(* IEC 61131-3 sources: plc-st-coding-agent/progress/evidence/f14_v10_full_20261113/jobs/codex_minimax-m27 (part 4) *)

(* ---- public-hard-06.raw_candidate_01.st ---- *)
(* ENGINEERING_CONTRACT *)
(*
┌──────────────────┬────────────────────────────────────────────────────────────────────────┐
│ Output/State     │ Activation, Retention, Reset, Priority, Units                          │
├──────────────────┼────────────────────────────────────────────────────────────────────────┤
│ MotorForward     │ Active during FEED, TRANSPORT_TO_WEIGH, TRANSPORT_TO_FIRING states     │
│                  │ in automatic mode only. Deactivated on state exit. PUB003, PUB006      │
├──────────────────┼────────────────────────────────────────────────────────────────────────┤
│ MotorReverse     │ Active during KICK state only (automatic mode). Deactivated on exit.   │
│                  │ Interlocked with MotorForward in manual mode. PUB002                   │
├──────────────────┼────────────────────────────────────────────────────────────────────────┤
│ kick             │ Latched HIGH when weight < 100 OR weight > 200 in WEIGH state.         │
│                  │ Deactivated when material exits wash station (SensorWash=FALSE).       │
│                  │ Single rejection per material cycle. PUB010                            │
├──────────────────┼────────────────────────────────────────────────────────────────────────┤
│ CompletionLight  │ Latched HIGH when SensorOutput=TRUE in OUTPUT state.                   │
│                  │ Deactivated when SensorOutput=FALSE (product removed).                 │
│                  │ No manual override specified. PUB012                                   │
├──────────────────┼────────────────────────────────────────────────────────────────────────┤
│ firingTemp       │ Calculated once when weight passes qualification check.                │
│                  │ Value: 500 + (weight - 100) * 0.5, range [500, 550]. Retained.         │
│                  │ PUB011                                                                   │
├──────────────────┼────────────────────────────────────────────────────────────────────────┤
│ State Machine    │ States: IDLE(0), FEED(1), WASH_WAIT(2), WEIGH(3), KICK(4),             │
│                  │ TRANSPORT_TO_FIRING(5), FIRING_WAIT(6), TRANSPORT_TO_OUTPUT(7),        │
│                  │ OUTPUT(8). Same-scan priority: sensor arrival > state transition.      │
│                  │ PUB003-PUB012                                                           │
└──────────────────┴────────────────────────────────────────────────────────────────────────┘
*)

(* CONTRACT_RULES [{"kind":"hold_until_reset","output":"CompletionLight","set_input":"SensorOutput","reset_input":"NOT SensorOutput"}] *)

FUNCTION_BLOCK ProductionControl
VAR
    tmp_state : INT := 0;
    tmp_prevSensorFeed : BOOL := FALSE;
    tmp_prevSensorWash : BOOL := FALSE;
    tmp_prevSensorWeight : BOOL := FALSE;
    tmp_prevSensorFiring : BOOL := FALSE;
END_VAR

// Reset all outputs at start of scan
MotorForward := FALSE;
MotorReverse := FALSE;
kick := FALSE;
CompletionLight := FALSE;

IF Mode = FALSE THEN
    // Manual Mode (PUB001, PUB002)
    MotorForward := ForwardButton AND NOT ReverseButton;
    MotorReverse := ReverseButton AND NOT ForwardButton;
ELSE
    // Automatic Mode (PUB003-PUB012)
    CASE tmp_state OF
        0: // IDLE - waiting for material at feed station
            IF SensorFeed THEN
                tmp_state := 1;
            END_IF;

        1: // FEED - transport to cleaning station
            MotorForward := TRUE;
            IF SensorWash THEN
                tmp_state := 2;
                MotorForward := FALSE;
            END_IF;

        2: // WASH_WAIT - waiting for cleaning completion
            IF washComplete THEN
                tmp_state := 3;
            END_IF;

        3: // WEIGH - process weight measurement
            IF weightComplete THEN
                IF weight < 100.0 OR weight > 200.0 THEN
                    // Unqualified: initiate kick
                    kick := TRUE;
                    MotorReverse := TRUE;
                    tmp_state := 4;
                ELSE
                    // Qualified: calculate firing temperature
                    firingTemp := 500.0 + (weight - 100.0) * 0.5;
                    MotorForward := TRUE;
                    tmp_state := 5;
                END_IF;
            END_IF;

        4: // KICK - reverse transport to exit wash station
            kick := TRUE;
            MotorReverse := TRUE;
            IF NOT SensorWash THEN
                kick := FALSE;
                MotorReverse := FALSE;
                tmp_state := 0;
            END_IF;

        5: // TRANSPORT_TO_FIRING
            MotorForward := TRUE;
            IF SensorFiring THEN
                tmp_state := 6;
                MotorForward := FALSE;
            END_IF;

        6: // FIRING_WAIT - waiting for firing completion
            IF firingComplete THEN
                tmp_state := 7;
            END_IF;

        7: // TRANSPORT_TO_OUTPUT
            MotorForward := TRUE;
            IF SensorOutput THEN
                tmp_state := 8;
                MotorForward := FALSE;
            END_IF;

        8: // OUTPUT - product complete, light on
            IF SensorOutput THEN
                CompletionLight := TRUE;
            ELSE
                CompletionLight := FALSE;
                tmp_state := 0;
            END_IF;

    END_CASE;
END_IF;

END_FUNCTION_BLOCK

(* ---- public-hard-06.raw_candidate_02.st ---- *)
(* ENGINEERING_CONTRACT *)
(*
┌──────────────────┬────────────────────────────────────────────────────────────────────────┐
│ Output/State     │ Activation, Retention, Reset, Priority, Units                          │
├──────────────────┼────────────────────────────────────────────────────────────────────────┤
│ MotorForward     │ Active during FEED, TRANSPORT_TO_WEIGH, TRANSPORT_TO_FIRING states     │
│                  │ in automatic mode only. Deactivated on state exit. PUB003, PUB006      │
├──────────────────┼────────────────────────────────────────────────────────────────────────┤
│ MotorReverse     │ Active during KICK state only (automatic mode). Deactivated on exit.   │
│                  │ Interlocked with MotorForward in manual mode. PUB002                   │
├──────────────────┼────────────────────────────────────────────────────────────────────────┤
│ kick             │ Latched HIGH when weight < 100 OR weight > 200 in WEIGH state.         │
│                  │ Deactivated when material exits wash station (SensorWash=FALSE).       │
│                  │ Single rejection per material cycle. PUB010                            │
├──────────────────┼────────────────────────────────────────────────────────────────────────┤
│ CompletionLight  │ Latched HIGH when SensorOutput=TRUE in OUTPUT state.                   │
│                  │ Deactivated when SensorOutput=FALSE (product removed).                 │
│                  │ No manual override specified. PUB012                                   │
├──────────────────┼────────────────────────────────────────────────────────────────────────┤
│ firingTemp       │ Calculated once when weight passes qualification check.                │
│                  │ Value: 500 + (weight - 100) * 0.5, range [500, 550]. Retained.         │
│                  │ PUB011                                                                   │
├──────────────────┼────────────────────────────────────────────────────────────────────────┤
│ State Machine    │ States: IDLE(0), FEED(1), WASH_WAIT(2), WEIGH(3), KICK(4),             │
│                  │ TRANSPORT_TO_FIRING(5), FIRING_WAIT(6), TRANSPORT_TO_OUTPUT(7),        │
│                  │ OUTPUT(8). Same-scan priority: sensor arrival > state transition.      │
│                  │ PUB003-PUB012                                                           │
└──────────────────┴────────────────────────────────────────────────────────────────────────┘
*)

(* CONTRACT_RULES [{"kind":"hold_until_reset","output":"CompletionLight","set_input":"SensorOutput","reset_input":"NOT SensorOutput"}] *)

FUNCTION_BLOCK ProductionControl
VAR_INPUT
    Mode : BOOL;
    ForwardButton : BOOL;
    ReverseButton : BOOL;
    SensorFeed : BOOL;
    SensorWash : BOOL;
    SensorWeight : BOOL;
    SensorFiring : BOOL;
    SensorOutput : BOOL;
    washComplete : BOOL;
    weightComplete : BOOL;
    weight : REAL;
    firingComplete : BOOL;
END_VAR

VAR_OUTPUT
    MotorForward : BOOL;
    MotorReverse : BOOL;
    kick : BOOL;
    CompletionLight : BOOL;
    firingTemp : REAL;
END_VAR

VAR
    tmp_state : INT := 0;
    tmp_prevSensorFeed : BOOL := FALSE;
    tmp_prevSensorWash : BOOL := FALSE;
    tmp_prevSensorWeight : BOOL := FALSE;
    tmp_prevSensorFiring : BOOL := FALSE;
END_VAR

// Reset all outputs at start of scan
MotorForward := FALSE;
MotorReverse := FALSE;
kick := FALSE;
CompletionLight := FALSE;

IF Mode = FALSE THEN
    // Manual Mode (PUB001, PUB002)
    MotorForward := ForwardButton AND NOT ReverseButton;
    MotorReverse := ReverseButton AND NOT ForwardButton;
ELSE
    // Automatic Mode (PUB003-PUB012)
    CASE tmp_state OF
        0: // IDLE - waiting for material at feed station
            IF SensorFeed THEN
                tmp_state := 1;
            END_IF;

        1: // FEED - transport to cleaning station
            MotorForward := TRUE;
            IF SensorWash THEN
                tmp_state := 2;
                MotorForward := FALSE;
            END_IF;

        2: // WASH_WAIT - waiting for cleaning completion
            IF washComplete THEN
                tmp_state := 3;
            END_IF;

        3: // WEIGH - process weight measurement
            IF weightComplete THEN
                IF weight < 100.0 OR weight > 200.0 THEN
                    // Unqualified: initiate kick
                    kick := TRUE;
                    MotorReverse := TRUE;
                    tmp_state := 4;
                ELSE
                    // Qualified: calculate firing temperature
                    firingTemp := 500.0 + (weight - 100.0) * 0.5;
                    MotorForward := TRUE;
                    tmp_state := 5;
                END_IF;
            END_IF;

        4: // KICK - reverse transport to exit wash station
            kick := TRUE;
            MotorReverse := TRUE;
            IF NOT SensorWash THEN
                kick := FALSE;
                MotorReverse := FALSE;
                tmp_state := 0;
            END_IF;

        5: // TRANSPORT_TO_FIRING
            MotorForward := TRUE;
            IF SensorFiring THEN
                tmp_state := 6;
                MotorForward := FALSE;
            END_IF;

        6: // FIRING_WAIT - waiting for firing completion
            IF firingComplete THEN
                tmp_state := 7;
            END_IF;

        7: // TRANSPORT_TO_OUTPUT
            MotorForward := TRUE;
            IF SensorOutput THEN
                tmp_state := 8;
                MotorForward := FALSE;
            END_IF;

        8: // OUTPUT - product complete, light on
            IF SensorOutput THEN
                CompletionLight := TRUE;
            ELSE
                CompletionLight := FALSE;
                tmp_state := 0;
            END_IF;

    END_CASE;
END_IF;

END_FUNCTION_BLOCK

(* ---- public-hard-06.raw_candidate_03.st ---- *)
(* ENGINEERING_CONTRACT *)
(*
┌──────────────────┬────────────────────────────────────────────────────────────────────────┐
│ Output/State     │ Activation, Retention, Reset, Priority, Units                          │
├──────────────────┼────────────────────────────────────────────────────────────────────────┤
│ MotorForward     │ Active during FEED, TRANSPORT_TO_WEIGH, TRANSPORT_TO_FIRING states     │
│                  │ in automatic mode only. Deactivated on state exit. PUB003, PUB006      │
├──────────────────┼────────────────────────────────────────────────────────────────────────┤
│ MotorReverse     │ Active during KICK state only (automatic mode). Deactivated on exit.   │
│                  │ Interlocked with MotorForward in manual mode. PUB002                   │
├──────────────────┼────────────────────────────────────────────────────────────────────────┤
│ kick             │ Latched HIGH when weight < 100 OR weight > 200 in WEIGH state.         │
│                  │ Deactivated when material exits wash station (SensorWash=FALSE).       │
│                  │ Single rejection per material cycle. PUB010                            │
├──────────────────┼────────────────────────────────────────────────────────────────────────┤
│ CompletionLight  │ Latched HIGH when SensorOutput=TRUE in OUTPUT state.                   │
│                  │ Deactivated when SensorOutput=FALSE (product removed).                 │
│                  │ No manual override specified. PUB012                                   │
├──────────────────┼────────────────────────────────────────────────────────────────────────┤
│ firingTemp       │ Calculated once when weight passes qualification check.                │
│                  │ Value: 500 + (weight - 100) * 0.5, range [500, 550]. Retained.         │
│                  │ PUB011                                                                   │
├──────────────────┼────────────────────────────────────────────────────────────────────────┤
│ State Machine    │ States: IDLE(0), FEED(1), WASH_WAIT(2), WEIGH(3), KICK(4),             │
│                  │ TRANSPORT_TO_FIRING(5), FIRING_WAIT(6), TRANSPORT_TO_OUTPUT(7),        │
│                  │ OUTPUT(8). Same-scan priority: sensor arrival > state transition.      │
│                  │ PUB003-PUB012                                                           │
└──────────────────┴────────────────────────────────────────────────────────────────────────┘
*)

(* CONTRACT_RULES [{"kind":"hold_until_reset","output":"CompletionLight","set_input":"SensorOutput","reset_input":"NOT SensorOutput"}] *)

FUNCTION_BLOCK ProductionControl
VAR_INPUT
    Mode : BOOL;
    ForwardButton : BOOL;
    ReverseButton : BOOL;
    SensorFeed : BOOL;
    SensorWash : BOOL;
    SensorWeight : BOOL;
    SensorFiring : BOOL;
    SensorOutput : BOOL;
    washComplete : BOOL;
    weightComplete : BOOL;
    weight : REAL;
    firingComplete : BOOL;
END_VAR

VAR_OUTPUT
    MotorForward : BOOL;
    MotorReverse : BOOL;
    kick : BOOL;
    CompletionLight : BOOL;
    firingTemp : REAL;
END_VAR

VAR
    tmp_state : INT := 0;
END_VAR

// Reset all outputs at start of scan
MotorForward := FALSE;
MotorReverse := FALSE;
kick := FALSE;
CompletionLight := FALSE;

IF Mode = FALSE THEN
    // Manual Mode (PUB001, PUB002)
    MotorForward := ForwardButton AND NOT ReverseButton;
    MotorReverse := ReverseButton AND NOT ForwardButton;
ELSE
    // Automatic Mode (PUB003-PUB012)
    CASE tmp_state OF
        0: // IDLE - waiting for material at feed station
            IF SensorFeed THEN
                tmp_state := 1;
                MotorForward := TRUE;
            END_IF;

        1: // FEED - transport to cleaning station
            MotorForward := TRUE;
            IF SensorWash THEN
                tmp_state := 2;
                MotorForward := FALSE;
            END_IF;

        2: // WASH_WAIT - waiting for cleaning completion
            IF washComplete THEN
                tmp_state := 3;
            END_IF;

        3: // WEIGH - process weight measurement
            IF weightComplete THEN
                IF weight < 100.0 OR weight > 200.0 THEN
                    // Unqualified: initiate kick
                    kick := TRUE;
                    MotorReverse := TRUE;
                    tmp_state := 4;
                ELSE
                    // Qualified: calculate firing temperature
                    firingTemp := 500.0 + (weight - 100.0) * 0.5;
                    MotorForward := TRUE;
                    tmp_state := 5;
                END_IF;
            END_IF;

        4: // KICK - reverse transport to exit wash station
            kick := TRUE;
            MotorReverse := TRUE;
            IF NOT SensorWash THEN
                kick := FALSE;
                MotorReverse := FALSE;
                tmp_state := 0;
            END_IF;

        5: // TRANSPORT_TO_FIRING
            MotorForward := TRUE;
            IF SensorFiring THEN
                tmp_state := 6;
                MotorForward := FALSE;
            END_IF;

        6: // FIRING_WAIT - waiting for firing completion
            IF firingComplete THEN
                tmp_state := 7;
            END_IF;

        7: // TRANSPORT_TO_OUTPUT
            MotorForward := TRUE;
            IF SensorOutput THEN
                tmp_state := 8;
                MotorForward := FALSE;
            END_IF;

        8: // OUTPUT - product complete, light on
            IF SensorOutput THEN
                CompletionLight := TRUE;
            ELSE
                CompletionLight := FALSE;
                tmp_state := 0;
            END_IF;

    END_CASE;
END_IF;

END_FUNCTION_BLOCK

(* ---- public-medium-01.candidate_01.st ---- *)
(* ENGINEERING_CONTRACT
===================
| Output/State        | Activation               | Retention | Explicit Reset | Same-Scan Priority | Units/Range |
|---------------------|--------------------------|-----------|----------------|--------------------|-------------|
| pumpGroup[].RunComd | start rising edge        | HOLD      | stop edge      | stop > start       | BOOL[1..5]  |
| Manual: selected    | selection=TRUE ∧ start   | HOLD      | stop edge      | stop > start       | pumpGroup   |
| Auto: top-3 priority| top-3 priority ∧ start   | HOLD      | stop edge      | stop > start       | sorted[1..3]|
| Mode switch         | immediate re-eval        | N/A       | N/A            | N/A                | mode BOOL   |

PUB001 (91-265): Mode determines Manual vs Auto selection logic
PUB002 (266-350): Manual mode uses pumpGroup[].selection as qualifier
PUB003 (351-463): Auto mode selects 3 highest-priority pumps
PUB004 (464-652): Stop button deactivates all pumps
*)
(* CONTRACT_RULES [] *)

FUNCTION_BLOCK FB_MultiPumpControl
VAR
    lastStart : BOOL := FALSE;
    lastStop  : BOOL := FALSE;
    stopped   : BOOL := FALSE;
    tmp_i     : INT;
    tmp_j     : INT;
    tmp_prio  : INT;
    tmp_sel   : BOOL;
    tmp_run   : BOOL;
END_VAR

tmp_sel := pumpGroup[1].selection; // Suppress unused warning

// Rising edge detection for stop
IF stop AND NOT lastStop THEN
    stopped := TRUE;
END_IF;

// Rising edge detection for start (only if not stopped)
IF start AND NOT lastStart AND NOT stopped THEN
    IF NOT mode THEN
        // Manual mode: start pumps where selection = TRUE
        FOR tmp_i := 1 TO 5 DO
            IF pumpGroup[tmp_i].selection THEN
                pumpGroup[tmp_i].RunComd := TRUE;
            END_IF;
        END_FOR;
    ELSE
        // Automatic mode: select top 3 by priority
        FOR tmp_i := 1 TO 4 DO
            FOR tmp_j := tmp_i + 1 TO 5 DO
                IF pumpGroup[tmp_j].priority > pumpGroup[tmp_i].priority THEN
                    tmp_prio := pumpGroup[tmp_i].priority;
                    tmp_sel  := pumpGroup[tmp_i].selection;
                    tmp_run  := pumpGroup[tmp_i].RunComd;

                    pumpGroup[tmp_i].priority := pumpGroup[tmp_j].priority;
                    pumpGroup[tmp_i].selection := pumpGroup[tmp_j].selection;
                    pumpGroup[tmp_i].RunComd   := pumpGroup[tmp_j].RunComd;

                    pumpGroup[tmp_j].priority := tmp_prio;
                    pumpGroup[tmp_j].selection := tmp_sel;
                    pumpGroup[tmp_j].RunComd   := tmp_run;
                END_IF;
            END_FOR;
        END_FOR;

        // Activate top 3 pumps (indices 1,2,3 after sort)
        FOR tmp_i := 1 TO 3 DO
            pumpGroup[tmp_i].RunComd := TRUE;
        END_FOR;
        FOR tmp_i := 4 TO 5 DO
            pumpGroup[tmp_i].RunComd := FALSE;
        END_FOR;
    END_IF;
END_IF;

// Rising edge detection for stop
IF stopped THEN
    FOR tmp_i := 1 TO 5 DO
        pumpGroup[tmp_i].RunComd := FALSE;
    END_FOR;
    stopped := FALSE;
END_IF;

lastStart := start;
lastStop  := stop;
END_FUNCTION_BLOCK

(* ---- public-medium-01.candidate_02.st ---- *)
(* ENGINEERING_CONTRACT
===================
| Output/State        | Activation               | Retention | Explicit Reset | Same-Scan Priority | Units/Range |
|---------------------|--------------------------|-----------|----------------|--------------------|-------------|
| pumpGroup[].RunComd | start rising edge        | HOLD      | stop edge      | stop > start       | BOOL[1..5]  |
| Manual: selected    | selection=TRUE ∧ start   | HOLD      | stop edge      | stop > start       | pumpGroup   |
| Auto: top-3 priority| top-3 priority ∧ start   | HOLD      | stop edge      | stop > start       | sorted[1..3]|
| Mode switch         | immediate re-eval        | N/A       | N/A            | N/A                | mode BOOL   |

PUB001 (91-265): Mode determines Manual vs Auto selection logic
PUB002 (266-350): Manual mode uses pumpGroup[].selection as qualifier
PUB003 (351-463): Auto mode selects 3 highest-priority pumps
PUB004 (464-652): Stop button deactivates all pumps
*)
(* CONTRACT_RULES [] *)

FUNCTION_BLOCK FB_MultiPumpControl
VAR_INPUT
    mode  : BOOL;
    start : BOOL;
    stop  : BOOL;
END_VAR
VAR_IN_OUT
    pumpGroup : ARRAY[1..5] OF ST_Pump;
END_VAR
VAR
    lastStart : BOOL := FALSE;
    lastStop  : BOOL := FALSE;
    startRising : BOOL := FALSE;
    stopRising  : BOOL := FALSE;
    tmp_i     : INT;
    tmp_j     : INT;
    tmp_prio  : INT;
    tmp_sel   : BOOL;
    tmp_run   : BOOL;
END_VAR

// Rising edge detection for start
startRising := start AND NOT lastStart;

// Rising edge detection for stop
stopRising := stop AND NOT lastStop;

// Rising edge: stop takes priority, stops all pumps immediately
IF stopRising THEN
    FOR tmp_i := 1 TO 5 DO
        pumpGroup[tmp_i].RunComd := FALSE;
    END_FOR;
END_IF;

// Rising edge: start activates pumps (only if stop not asserted this scan)
IF startRising AND NOT stopRising THEN
    IF NOT mode THEN
        // Manual mode: start pumps where selection = TRUE
        FOR tmp_i := 1 TO 5 DO
            IF pumpGroup[tmp_i].selection THEN
                pumpGroup[tmp_i].RunComd := TRUE;
            END_IF;
        END_FOR;
    ELSE
        // Automatic mode: select top 3 by priority (bubble sort descending)
        FOR tmp_i := 1 TO 4 DO
            FOR tmp_j := tmp_i + 1 TO 5 DO
                IF pumpGroup[tmp_j].priority > pumpGroup[tmp_i].priority THEN
                    tmp_prio := pumpGroup[tmp_i].priority;
                    tmp_sel  := pumpGroup[tmp_i].selection;
                    tmp_run  := pumpGroup[tmp_i].RunComd;

                    pumpGroup[tmp_i].priority := pumpGroup[tmp_j].priority;
                    pumpGroup[tmp_i].selection := pumpGroup[tmp_j].selection;
                    pumpGroup[tmp_i].RunComd   := pumpGroup[tmp_j].RunComd;

                    pumpGroup[tmp_j].priority := tmp_prio;
                    pumpGroup[tmp_j].selection := tmp_sel;
                    pumpGroup[tmp_j].RunComd   := tmp_run;
                END_IF;
            END_FOR;
        END_FOR;

        // Activate top 3 pumps (indices 1,2,3 after sort)
        FOR tmp_i := 1 TO 3 DO
            pumpGroup[tmp_i].RunComd := TRUE;
        END_FOR;
        // Deactivate remaining pumps
        FOR tmp_i := 4 TO 5 DO
            pumpGroup[tmp_i].RunComd := FALSE;
        END_FOR;
    END_IF;
END_IF;

lastStart := start;
lastStop  := stop;
END_FUNCTION_BLOCK

(* ---- public-medium-01.candidate_03.st ---- *)
FUNCTION_BLOCK FB_MultiPumpControl
VAR_INPUT
    mode  : BOOL;
    start : BOOL;
    stop  : BOOL;
END_VAR

VAR_IN_OUT
    pumpGroup : ARRAY[1..5] OF ST_Pump;
END_VAR

VAR
    lastStart : BOOL := FALSE;
    lastStop  : BOOL := FALSE;
    stopped   : BOOL := FALSE;
    tmp_i     : INT;
    tmp_j     : INT;
    tmp_prio  : INT;
    tmp_sel   : BOOL;
    tmp_run   : BOOL;
END_VAR

// Rising edge detection for stop
IF stop AND NOT lastStop THEN
    stopped := TRUE;
END_IF;

// Rising edge detection for start (only if not stopped)
IF start AND NOT lastStart AND NOT stopped THEN
    IF NOT mode THEN
        // Manual mode: start pumps where selection = TRUE
        FOR tmp_i := 1 TO 5 DO
            IF pumpGroup[tmp_i].selection THEN
                pumpGroup[tmp_i].RunComd := TRUE;
            END_IF;
        END_FOR;
    ELSE
        // Automatic mode: select top 3 by priority
        FOR tmp_i := 1 TO 4 DO
            FOR tmp_j := tmp_i + 1 TO 5 DO
                IF pumpGroup[tmp_j].priority > pumpGroup[tmp_i].priority THEN
                    tmp_prio := pumpGroup[tmp_i].priority;
                    tmp_sel  := pumpGroup[tmp_i].selection;
                    tmp_run  := pumpGroup[tmp_i].RunComd;

                    pumpGroup[tmp_i].priority := pumpGroup[tmp_j].priority;
                    pumpGroup[tmp_i].selection := pumpGroup[tmp_j].selection;
                    pumpGroup[tmp_i].RunComd   := pumpGroup[tmp_j].RunComd;

                    pumpGroup[tmp_j].priority := tmp_prio;
                    pumpGroup[tmp_j].selection := tmp_sel;
                    pumpGroup[tmp_j].RunComd   := tmp_run;
                END_IF;
            END_FOR;
        END_FOR;

        // Activate top 3 pumps (indices 1,2,3 after sort)
        FOR tmp_i := 1 TO 3 DO
            pumpGroup[tmp_i].RunComd := TRUE;
        END_FOR;
        FOR tmp_i := 4 TO 5 DO
            pumpGroup[tmp_i].RunComd := FALSE;
        END_FOR;
    END_IF;
END_IF;

// Rising edge detection for stop
IF stopped THEN
    FOR tmp_i := 1 TO 5 DO
        pumpGroup[tmp_i].RunComd := FALSE;
    END_FOR;
    stopped := FALSE;
END_IF;

lastStart := start;
lastStop  := stop;
END_FUNCTION_BLOCK

(* ---- public-medium-01.candidate_04.st ---- *)
Looking at the compilation errors, the main issues are:
1. Missing `FUNCTION_BLOCK` declaration line
2. Missing `VAR_INPUT` section for `mode`, `start`, `stop`
3. Missing `VAR_IN_OUT` section for `pumpGroup`
4. The `tmp_sel` assignment line needs proper structure access

(* ENGINEERING_CONTRACT
===================
| Output/State        | Activation               | Retention | Explicit Reset | Same-Scan Priority | Units/Range |
|---------------------|--------------------------|-----------|----------------|--------------------|-------------|
| pumpGroup[].RunComd | start rising edge        | HOLD      | stop edge      | stop > start       | BOOL[1..5]  |
| Manual: selected    | selection=TRUE ∧ start   | HOLD      | stop edge      | stop > start       | pumpGroup   |
| Auto: top-3 priority| top-3 priority ∧ start   | HOLD      | stop edge      | stop > start       | sorted[1..3]|
| Mode switch         | immediate re-eval        | N/A       | N/A            | N/A                | mode BOOL   |

PUB001 (91-265): Mode determines Manual vs Auto selection logic
PUB002 (266-350): Manual mode uses pumpGroup[].selection as qualifier
PUB003 (351-463): Auto mode selects 3 highest-priority pumps
PUB004 (464-652): Stop button deactivates all pumps
*)
(* CONTRACT_RULES [] *)

FUNCTION_BLOCK FB_MultiPumpControl
VAR_INPUT
    mode  : BOOL;
    start : BOOL;
    stop  : BOOL;
END_VAR
VAR_IN_OUT
    pumpGroup : ARRAY[1..5] OF ST_Pump;
END_VAR
VAR
    lastStart : BOOL := FALSE;
    lastStop  : BOOL := FALSE;
    stopped   : BOOL := FALSE;
    tmp_i     : INT;
    tmp_j     : INT;
    tmp_prio  : INT;
    tmp_sel   : BOOL;
    tmp_run   : BOOL;
END_VAR

tmp_sel := pumpGroup[1].selection;

IF stop AND NOT lastStop THEN
    stopped := TRUE;
END_IF;

IF start AND NOT lastStart AND NOT stopped THEN
    IF NOT mode THEN
        FOR tmp_i := 1 TO 5 DO
            IF pumpGroup[tmp_i].selection THEN
                pumpGroup[tmp_i].RunComd := TRUE;
            END_IF;
        END_FOR;
    ELSE
        FOR tmp_i := 1 TO 4 DO
            FOR tmp_j := tmp_i + 1 TO 5 DO
                IF pumpGroup[tmp_j].priority > pumpGroup[tmp_i].priority THEN
                    tmp_prio := pumpGroup[tmp_i].priority;
                    tmp_sel  := pumpGroup[tmp_i].selection;
                    tmp_run  := pumpGroup[tmp_i].RunComd;

                    pumpGroup[tmp_i].priority := pumpGroup[tmp_j].priority;
                    pumpGroup[tmp_i].selection := pumpGroup[tmp_j].selection;
                    pumpGroup[tmp_i].RunComd   := pumpGroup[tmp_j].RunComd;

                    pumpGroup[tmp_j].priority := tmp_prio;
                    pumpGroup[tmp_j].selection := tmp_sel;
                    pumpGroup[tmp_j].RunComd   := tmp_run;
                END_IF;
            END_FOR;
        END_FOR;

        FOR tmp_i := 1 TO 3 DO
            pumpGroup[tmp_i].RunComd := TRUE;
        END_FOR;
        FOR tmp_i := 4 TO 5 DO
            pumpGroup[tmp_i].RunComd := FALSE;
        END_FOR;
    END_IF;
END_IF;

IF stopped THEN
    FOR tmp_i := 1 TO 5 DO
        pumpGroup[tmp_i].RunComd := FALSE;
    END_FOR;
    stopped := FALSE;
END_IF;

lastStart := start;
lastStop  := stop;
END_FUNCTION_BLOCK

(* ---- public-medium-01.raw_candidate_01.st ---- *)
(* ENGINEERING_CONTRACT
===================
| Output/State        | Activation               | Retention | Explicit Reset | Same-Scan Priority | Units/Range |
|---------------------|--------------------------|-----------|----------------|--------------------|-------------|
| pumpGroup[].RunComd | start rising edge        | HOLD      | stop edge      | stop > start       | BOOL[1..5]  |
| Manual: selected    | selection=TRUE ∧ start   | HOLD      | stop edge      | stop > start       | pumpGroup   |
| Auto: top-3 priority| top-3 priority ∧ start   | HOLD      | stop edge      | stop > start       | sorted[1..3]|
| Mode switch         | immediate re-eval        | N/A       | N/A            | N/A                | mode BOOL   |

PUB001 (91-265): Mode determines Manual vs Auto selection logic
PUB002 (266-350): Manual mode uses pumpGroup[].selection as qualifier
PUB003 (351-463): Auto mode selects 3 highest-priority pumps
PUB004 (464-652): Stop button deactivates all pumps
*)
(* CONTRACT_RULES [] *)

FUNCTION_BLOCK FB_MultiPumpControl
VAR
    lastStart : BOOL := FALSE;
    lastStop  : BOOL := FALSE;
    stopped   : BOOL := FALSE;
    tmp_i     : INT;
    tmp_j     : INT;
    tmp_prio  : INT;
    tmp_sel   : BOOL;
    tmp_run   : BOOL;
END_VAR

tmp_sel := pumpGroup[1].selection; // Suppress unused warning

// Rising edge detection for stop
IF stop AND NOT lastStop THEN
    stopped := TRUE;
END_IF;

// Rising edge detection for start (only if not stopped)
IF start AND NOT lastStart AND NOT stopped THEN
    IF NOT mode THEN
        // Manual mode: start pumps where selection = TRUE
        FOR tmp_i := 1 TO 5 DO
            IF pumpGroup[tmp_i].selection THEN
                pumpGroup[tmp_i].RunComd := TRUE;
            END_IF;
        END_FOR;
    ELSE
        // Automatic mode: select top 3 by priority
        FOR tmp_i := 1 TO 4 DO
            FOR tmp_j := tmp_i + 1 TO 5 DO
                IF pumpGroup[tmp_j].priority > pumpGroup[tmp_i].priority THEN
                    tmp_prio := pumpGroup[tmp_i].priority;
                    tmp_sel  := pumpGroup[tmp_i].selection;
                    tmp_run  := pumpGroup[tmp_i].RunComd;

                    pumpGroup[tmp_i].priority := pumpGroup[tmp_j].priority;
                    pumpGroup[tmp_i].selection := pumpGroup[tmp_j].selection;
                    pumpGroup[tmp_i].RunComd   := pumpGroup[tmp_j].RunComd;

                    pumpGroup[tmp_j].priority := tmp_prio;
                    pumpGroup[tmp_j].selection := tmp_sel;
                    pumpGroup[tmp_j].RunComd   := tmp_run;
                END_IF;
            END_FOR;
        END_FOR;

        // Activate top 3 pumps (indices 1,2,3 after sort)
        FOR tmp_i := 1 TO 3 DO
            pumpGroup[tmp_i].RunComd := TRUE;
        END_FOR;
        FOR tmp_i := 4 TO 5 DO
            pumpGroup[tmp_i].RunComd := FALSE;
        END_FOR;
    END_IF;
END_IF;

// Rising edge detection for stop
IF stopped THEN
    FOR tmp_i := 1 TO 5 DO
        pumpGroup[tmp_i].RunComd := FALSE;
    END_FOR;
    stopped := FALSE;
END_IF;

lastStart := start;
lastStop  := stop;
END_FUNCTION_BLOCK

(* ---- public-medium-01.raw_candidate_02.st ---- *)
(* ENGINEERING_CONTRACT
===================
| Output/State        | Activation               | Retention | Explicit Reset | Same-Scan Priority | Units/Range |
|---------------------|--------------------------|-----------|----------------|--------------------|-------------|
| pumpGroup[].RunComd | start rising edge        | HOLD      | stop edge      | stop > start       | BOOL[1..5]  |
| Manual: selected    | selection=TRUE ∧ start   | HOLD      | stop edge      | stop > start       | pumpGroup   |
| Auto: top-3 priority| top-3 priority ∧ start   | HOLD      | stop edge      | stop > start       | sorted[1..3]|
| Mode switch         | immediate re-eval        | N/A       | N/A            | N/A                | mode BOOL   |

PUB001 (91-265): Mode determines Manual vs Auto selection logic
PUB002 (266-350): Manual mode uses pumpGroup[].selection as qualifier
PUB003 (351-463): Auto mode selects 3 highest-priority pumps
PUB004 (464-652): Stop button deactivates all pumps
*)
(* CONTRACT_RULES [] *)

FUNCTION_BLOCK FB_MultiPumpControl
VAR_INPUT
    mode  : BOOL;
    start : BOOL;
    stop  : BOOL;
END_VAR
VAR_IN_OUT
    pumpGroup : ARRAY[1..5] OF ST_Pump;
END_VAR
VAR
    lastStart : BOOL := FALSE;
    lastStop  : BOOL := FALSE;
    startRising : BOOL := FALSE;
    stopRising  : BOOL := FALSE;
    tmp_i     : INT;
    tmp_j     : INT;
    tmp_prio  : INT;
    tmp_sel   : BOOL;
    tmp_run   : BOOL;
END_VAR

// Rising edge detection for start
startRising := start AND NOT lastStart;

// Rising edge detection for stop
stopRising := stop AND NOT lastStop;

// Rising edge: stop takes priority, stops all pumps immediately
IF stopRising THEN
    FOR tmp_i := 1 TO 5 DO
        pumpGroup[tmp_i].RunComd := FALSE;
    END_FOR;
END_IF;

// Rising edge: start activates pumps (only if stop not asserted this scan)
IF startRising AND NOT stopRising THEN
    IF NOT mode THEN
        // Manual mode: start pumps where selection = TRUE
        FOR tmp_i := 1 TO 5 DO
            IF pumpGroup[tmp_i].selection THEN
                pumpGroup[tmp_i].RunComd := TRUE;
            END_IF;
        END_FOR;
    ELSE
        // Automatic mode: select top 3 by priority (bubble sort descending)
        FOR tmp_i := 1 TO 4 DO
            FOR tmp_j := tmp_i + 1 TO 5 DO
                IF pumpGroup[tmp_j].priority > pumpGroup[tmp_i].priority THEN
                    tmp_prio := pumpGroup[tmp_i].priority;
                    tmp_sel  := pumpGroup[tmp_i].selection;
                    tmp_run  := pumpGroup[tmp_i].RunComd;

                    pumpGroup[tmp_i].priority := pumpGroup[tmp_j].priority;
                    pumpGroup[tmp_i].selection := pumpGroup[tmp_j].selection;
                    pumpGroup[tmp_i].RunComd   := pumpGroup[tmp_j].RunComd;

                    pumpGroup[tmp_j].priority := tmp_prio;
                    pumpGroup[tmp_j].selection := tmp_sel;
                    pumpGroup[tmp_j].RunComd   := tmp_run;
                END_IF;
            END_FOR;
        END_FOR;

        // Activate top 3 pumps (indices 1,2,3 after sort)
        FOR tmp_i := 1 TO 3 DO
            pumpGroup[tmp_i].RunComd := TRUE;
        END_FOR;
        // Deactivate remaining pumps
        FOR tmp_i := 4 TO 5 DO
            pumpGroup[tmp_i].RunComd := FALSE;
        END_FOR;
    END_IF;
END_IF;

lastStart := start;
lastStop  := stop;
END_FUNCTION_BLOCK

(* ---- public-medium-01.raw_candidate_03.st ---- *)
FUNCTION_BLOCK FB_MultiPumpControl
VAR_INPUT
    mode  : BOOL;
    start : BOOL;
    stop  : BOOL;
END_VAR

VAR_IN_OUT
    pumpGroup : ARRAY[1..5] OF ST_Pump;
END_VAR

VAR
    lastStart : BOOL := FALSE;
    lastStop  : BOOL := FALSE;
    stopped   : BOOL := FALSE;
    tmp_i     : INT;
    tmp_j     : INT;
    tmp_prio  : INT;
    tmp_sel   : BOOL;
    tmp_run   : BOOL;
END_VAR

// Rising edge detection for stop
IF stop AND NOT lastStop THEN
    stopped := TRUE;
END_IF;

// Rising edge detection for start (only if not stopped)
IF start AND NOT lastStart AND NOT stopped THEN
    IF NOT mode THEN
        // Manual mode: start pumps where selection = TRUE
        FOR tmp_i := 1 TO 5 DO
            IF pumpGroup[tmp_i].selection THEN
                pumpGroup[tmp_i].RunComd := TRUE;
            END_IF;
        END_FOR;
    ELSE
        // Automatic mode: select top 3 by priority
        FOR tmp_i := 1 TO 4 DO
            FOR tmp_j := tmp_i + 1 TO 5 DO
                IF pumpGroup[tmp_j].priority > pumpGroup[tmp_i].priority THEN
                    tmp_prio := pumpGroup[tmp_i].priority;
                    tmp_sel  := pumpGroup[tmp_i].selection;
                    tmp_run  := pumpGroup[tmp_i].RunComd;

                    pumpGroup[tmp_i].priority := pumpGroup[tmp_j].priority;
                    pumpGroup[tmp_i].selection := pumpGroup[tmp_j].selection;
                    pumpGroup[tmp_i].RunComd   := pumpGroup[tmp_j].RunComd;

                    pumpGroup[tmp_j].priority := tmp_prio;
                    pumpGroup[tmp_j].selection := tmp_sel;
                    pumpGroup[tmp_j].RunComd   := tmp_run;
                END_IF;
            END_FOR;
        END_FOR;

        // Activate top 3 pumps (indices 1,2,3 after sort)
        FOR tmp_i := 1 TO 3 DO
            pumpGroup[tmp_i].RunComd := TRUE;
        END_FOR;
        FOR tmp_i := 4 TO 5 DO
            pumpGroup[tmp_i].RunComd := FALSE;
        END_FOR;
    END_IF;
END_IF;

// Rising edge detection for stop
IF stopped THEN
    FOR tmp_i := 1 TO 5 DO
        pumpGroup[tmp_i].RunComd := FALSE;
    END_FOR;
    stopped := FALSE;
END_IF;

lastStart := start;
lastStop  := stop;
END_FUNCTION_BLOCK

(* ---- public-medium-01.raw_candidate_04.st ---- *)
Looking at the compilation errors, the main issues are:
1. Missing `FUNCTION_BLOCK` declaration line
2. Missing `VAR_INPUT` section for `mode`, `start`, `stop`
3. Missing `VAR_IN_OUT` section for `pumpGroup`
4. The `tmp_sel` assignment line needs proper structure access

(* ENGINEERING_CONTRACT
===================
| Output/State        | Activation               | Retention | Explicit Reset | Same-Scan Priority | Units/Range |
|---------------------|--------------------------|-----------|----------------|--------------------|-------------|
| pumpGroup[].RunComd | start rising edge        | HOLD      | stop edge      | stop > start       | BOOL[1..5]  |
| Manual: selected    | selection=TRUE ∧ start   | HOLD      | stop edge      | stop > start       | pumpGroup   |
| Auto: top-3 priority| top-3 priority ∧ start   | HOLD      | stop edge      | stop > start       | sorted[1..3]|
| Mode switch         | immediate re-eval        | N/A       | N/A            | N/A                | mode BOOL   |

PUB001 (91-265): Mode determines Manual vs Auto selection logic
PUB002 (266-350): Manual mode uses pumpGroup[].selection as qualifier
PUB003 (351-463): Auto mode selects 3 highest-priority pumps
PUB004 (464-652): Stop button deactivates all pumps
*)
(* CONTRACT_RULES [] *)

FUNCTION_BLOCK FB_MultiPumpControl
VAR_INPUT
    mode  : BOOL;
    start : BOOL;
    stop  : BOOL;
END_VAR
VAR_IN_OUT
    pumpGroup : ARRAY[1..5] OF ST_Pump;
END_VAR
VAR
    lastStart : BOOL := FALSE;
    lastStop  : BOOL := FALSE;
    stopped   : BOOL := FALSE;
    tmp_i     : INT;
    tmp_j     : INT;
    tmp_prio  : INT;
    tmp_sel   : BOOL;
    tmp_run   : BOOL;
END_VAR

tmp_sel := pumpGroup[1].selection;

IF stop AND NOT lastStop THEN
    stopped := TRUE;
END_IF;

IF start AND NOT lastStart AND NOT stopped THEN
    IF NOT mode THEN
        FOR tmp_i := 1 TO 5 DO
            IF pumpGroup[tmp_i].selection THEN
                pumpGroup[tmp_i].RunComd := TRUE;
            END_IF;
        END_FOR;
    ELSE
        FOR tmp_i := 1 TO 4 DO
            FOR tmp_j := tmp_i + 1 TO 5 DO
                IF pumpGroup[tmp_j].priority > pumpGroup[tmp_i].priority THEN
                    tmp_prio := pumpGroup[tmp_i].priority;
                    tmp_sel  := pumpGroup[tmp_i].selection;
                    tmp_run  := pumpGroup[tmp_i].RunComd;

                    pumpGroup[tmp_i].priority := pumpGroup[tmp_j].priority;
                    pumpGroup[tmp_i].selection := pumpGroup[tmp_j].selection;
                    pumpGroup[tmp_i].RunComd   := pumpGroup[tmp_j].RunComd;

                    pumpGroup[tmp_j].priority := tmp_prio;
                    pumpGroup[tmp_j].selection := tmp_sel;
                    pumpGroup[tmp_j].RunComd   := tmp_run;
                END_IF;
            END_FOR;
        END_FOR;

        FOR tmp_i := 1 TO 3 DO
            pumpGroup[tmp_i].RunComd := TRUE;
        END_FOR;
        FOR tmp_i := 4 TO 5 DO
            pumpGroup[tmp_i].RunComd := FALSE;
        END_FOR;
    END_IF;
END_IF;

IF stopped THEN
    FOR tmp_i := 1 TO 5 DO
        pumpGroup[tmp_i].RunComd := FALSE;
    END_FOR;
    stopped := FALSE;
END_IF;

lastStart := start;
lastStop  := stop;
END_FUNCTION_BLOCK

(* ---- public-medium-02.candidate_01.st ---- *)
FUNCTION_BLOCK AnalogBatchProcessing
VAR_INPUT
    count : DINT;
END_VAR
VAR_IN_OUT
    analogValues : ARRAY[*] OF INT;
    channels     : ARRAY[*] OF ST_AnalogChannel;
END_VAR
VAR
    tmp_i         : DINT;
    tmp_rawMin    : REAL;
    tmp_rawMax    : REAL;
    tmp_rawRange  : REAL;
    tmp_engRange  : REAL;
    tmp_raw       : INT;
    tmp_analogVal : REAL;
END_VAR
(* CONTRACT_RULES [] *)
(* ENGINEERING_CONTRACT
 * Activation:       Each scan processes up to 'count' channels sequentially.
 * Retention:        retVal and outputValue are overwritten each scan; no latching.
 * Explicit Reset:   None specified; outputs refresh every scan.
 * Same-scan Priority: Sequential ordinal processing; first failure does not halt loop.
 * Units/Boundaries:
 *   - PUB001: count is caller-supplied bound selector; arrays use their own lower bounds.
 *   - PUB002: measuringMode 0=linear (bipolar/unipolar), 1=std temp (÷10), 2=climatic (÷100).
 *   - PUB003: Linear scaling uses full-scale raw range; output = loLIM + ratio*(hiLIM-loLIM).
 *   - PUB004: RetVal 16#8001 on invalid measuringMode; 16#8002 on hiLIM<=loLIM.
 *   - PUB005: OutputValue written only on successful conversion; retVal set on error.
 *   - PUB006: Disabled channels (enable=FALSE) are skipped without modifying retVal/outputValue.
 *   - PUB007: All arithmetic uses REAL; explicit conversions applied to raw INT operands.
 *   - PUB008: No delay, no edge detection, no state machine; pure per-scan calculation.
 *)

    tmp_i := LOWER_BOUND(analogValues, 1);

    WHILE tmp_i < LOWER_BOUND(analogValues, 1) + count DO
        IF channels[tmp_i].enable THEN
            IF channels[tmp_i].hiLIM <= channels[tmp_i].loLIM THEN
                channels[tmp_i].retVal := 16#8002;
            ELSE
                CASE channels[tmp_i].measuringMode OF
                    0: // Non-temperature linear scaling
                        tmp_raw := analogValues[tmp_i];
                        tmp_analogVal := TO_REAL(tmp_raw);

                        IF channels[tmp_i].bipolar THEN
                            tmp_rawMin := TO_REAL(-27648);
                            tmp_rawMax := TO_REAL(27648);
                        ELSE
                            tmp_rawMin := TO_REAL(0);
                            tmp_rawMax := TO_REAL(27648);
                        END_IF;

                        tmp_rawRange := tmp_rawMax - tmp_rawMin;
                        tmp_engRange := channels[tmp_i].hiLIM - channels[tmp_i].loLIM;

                        channels[tmp_i].outputValue := channels[tmp_i].loLIM +
                            ((tmp_analogVal - tmp_rawMin) / tmp_rawRange) * tmp_engRange;
                        channels[tmp_i].retVal := 16#0000;

                    1: // Standard temperature
                        tmp_raw := analogValues[tmp_i];
                        channels[tmp_i].outputValue := TO_REAL(tmp_raw) / 10.0;
                        channels[tmp_i].retVal := 16#0000;

                    2: // Climatic temperature
                        tmp_raw := analogValues[tmp_i];
                        channels[tmp_i].outputValue := TO_REAL(tmp_raw) / 100.0;
                        channels[tmp_i].retVal := 16#0000;

                    ELSE
                        channels[tmp_i].retVal := 16#8001;
                END_CASE;
            END_IF;
        END_IF;

        tmp_i := tmp_i + 1;
    END_WHILE;

END_FUNCTION_BLOCK

(* ---- public-medium-02.candidate_02.st ---- *)
TYPE ST_AnalogChannel :
STRUCT
    enable        : BOOL;
    hiLIM         : REAL;
    loLIM         : REAL;
    bipolar       : BOOL;
    measuringMode : INT;
    retVal        : WORD;
    outputValue   : REAL;
END_STRUCT
END_TYPE;

FUNCTION_BLOCK AnalogBatchProcessing
VAR_INPUT
    count : DINT;
END_VAR
VAR_IN_OUT
    analogValues : ARRAY[*] OF INT;
    channels     : ARRAY[*] OF ST_AnalogChannel;
END_VAR
VAR
    tmp_i         : DINT;
    tmp_rawMin    : REAL;
    tmp_rawMax    : REAL;
    tmp_rawRange  : REAL;
    tmp_engRange  : REAL;
    tmp_raw       : INT;
    tmp_analogVal : REAL;
END_VAR
(* CONTRACT_RULES [] *)
(* ENGINEERING_CONTRACT
 * Activation:       Each scan processes up to 'count' channels sequentially.
 * Retention:        retVal and outputValue are overwritten each scan; no latching.
 * Explicit Reset:   None specified; outputs refresh every scan.
 * Same-scan Priority: Sequential ordinal processing; first failure does not halt loop.
 * Units/Boundaries:
 *   - PUB001: count is caller-supplied bound selector; arrays use their own lower bounds.
 *   - PUB002: measuringMode 0=linear (bipolar/unipolar), 1=std temp (÷10), 2=climatic (÷100).
 *   - PUB003: Linear scaling uses full-scale raw range; output = loLIM + ratio*(hiLIM-loLIM).
 *   - PUB004: RetVal 16#8001 on invalid measuringMode; 16#8002 on hiLIM<=loLIM.
 *   - PUB005: OutputValue written only on successful conversion; retVal set on error.
 *   - PUB006: Disabled channels (enable=FALSE) are skipped without modifying retVal/outputValue.
 *   - PUB007: All arithmetic uses REAL; explicit conversions applied to raw INT operands.
 *   - PUB008: No delay, no edge detection, no state machine; pure per-scan calculation.
 *)

    tmp_i := LOWER_BOUND(analogValues, 1);

    WHILE tmp_i < LOWER_BOUND(analogValues, 1) + count DO
        IF channels[tmp_i].enable THEN
            IF channels[tmp_i].hiLIM <= channels[tmp_i].loLIM THEN
                channels[tmp_i].retVal := 16#8002;
            ELSE
                CASE channels[tmp_i].measuringMode OF
                    0: // Non-temperature linear scaling
                        tmp_raw := analogValues[tmp_i];
                        tmp_analogVal := TO_REAL(tmp_raw);

                        IF channels[tmp_i].bipolar THEN
                            tmp_rawMin := TO_REAL(-27648);
                            tmp_rawMax := TO_REAL(27648);
                        ELSE
                            tmp_rawMin := TO_REAL(0);
                            tmp_rawMax := TO_REAL(27648);
                        END_IF;

                        tmp_rawRange := tmp_rawMax - tmp_rawMin;
                        tmp_engRange := channels[tmp_i].hiLIM - channels[tmp_i].loLIM;

                        channels[tmp_i].outputValue := channels[tmp_i].loLIM +
                            ((tmp_analogVal - tmp_rawMin) / tmp_rawRange) * tmp_engRange;
                        channels[tmp_i].retVal := 16#0000;

                    1: // Standard temperature
                        tmp_raw := analogValues[tmp_i];
                        channels[tmp_i].outputValue := TO_REAL(tmp_raw) / 10.0;
                        channels[tmp_i].retVal := 16#0000;

                    2: // Climatic temperature
                        tmp_raw := analogValues[tmp_i];
                        channels[tmp_i].outputValue := TO_REAL(tmp_raw) / 100.0;
                        channels[tmp_i].retVal := 16#0000;

                    ELSE
                        channels[tmp_i].retVal := 16#8001;
                END_CASE;
            END_IF;
        END_IF;

        tmp_i := tmp_i + 1;
    END_WHILE;

END_FUNCTION_BLOCK

(* ---- public-medium-02.candidate_03.st ---- *)
TYPE ST_AnalogChannel :
STRUCT
    enable        : BOOL;
    hiLIM         : REAL;
    loLIM         : REAL;
    bipolar       : BOOL;
    measuringMode : INT;
    retVal        : WORD;
    outputValue   : REAL;
END_STRUCT
END_TYPE;

FUNCTION_BLOCK AnalogBatchProcessing
VAR_INPUT
    count : DINT;
END_VAR
VAR_IN_OUT
    analogValues : ARRAY[*] OF INT;
    channels     : ARRAY[*] OF ST_AnalogChannel;
END_VAR
VAR
    tmp_i             : DINT;
    tmp_channelsLower : DINT;
    tmp_analogLower   : DINT;
    tmp_rawMin        : REAL;
    tmp_rawMax        : REAL;
    tmp_rawRange      : REAL;
    tmp_engRange      : REAL;
    tmp_raw           : INT;
    tmp_analogVal     : REAL;
END_VAR
(* CONTRACT_RULES [] *)
(* ENGINEERING_CONTRACT
 * Activation:       Each scan processes up to 'count' channels sequentially.
 * Retention:        retVal and outputValue are overwritten each scan; no latching.
 * Explicit Reset:   None specified; outputs refresh every scan.
 * Same-scan Priority: Sequential ordinal processing; first failure does not halt loop.
 * Units/Boundaries:
 *   - PUB001: count is caller-supplied bound selector; arrays use their own lower bounds.
 *   - PUB002: measuringMode 0=linear (bipolar/unipolar), 1=std temp (÷10), 2=climatic (÷100).
 *   - PUB003: Linear scaling uses full-scale raw range; output = loLIM + ratio*(hiLIM-loLIM).
 *   - PUB004: RetVal 16#8001 on invalid measuringMode; 16#8002 on hiLIM<=loLIM.
 *   - PUB005: OutputValue written only on successful conversion; retVal set on error.
 *   - PUB006: Disabled channels (enable=FALSE) are skipped without modifying retVal/outputValue.
 *   - PUB007: All arithmetic uses REAL; explicit conversions applied to raw INT operands.
 *   - PUB008: No delay, no edge detection, no state machine; pure per-scan calculation.
 *)

    tmp_channelsLower := LOWER_BOUND(channels, 1);
    tmp_analogLower   := LOWER_BOUND(analogValues, 1);
    tmp_i := tmp_channelsLower;

    WHILE tmp_i < tmp_channelsLower + count DO
        IF channels[tmp_i].enable THEN
            IF channels[tmp_i].hiLIM <= channels[tmp_i].loLIM THEN
                channels[tmp_i].retVal := 16#8002;
            ELSE
                CASE channels[tmp_i].measuringMode OF
                    0: // Non-temperature linear scaling
                        tmp_raw := analogValues[tmp_analogLower + (tmp_i - tmp_channelsLower)];
                        tmp_analogVal := TO_REAL(tmp_raw);

                        IF channels[tmp_i].bipolar THEN
                            tmp_rawMin := TO_REAL(-27648);
                            tmp_rawMax := TO_REAL(27648);
                        ELSE
                            tmp_rawMin := TO_REAL(0);
                            tmp_rawMax := TO_REAL(27648);
                        END_IF;

                        tmp_rawRange := tmp_rawMax - tmp_rawMin;
                        tmp_engRange := channels[tmp_i].hiLIM - channels[tmp_i].loLIM;

                        channels[tmp_i].outputValue := channels[tmp_i].loLIM +
                            ((tmp_analogVal - tmp_rawMin) / tmp_rawRange) * tmp_engRange;
                        channels[tmp_i].retVal := 16#0000;

                    1: // Standard temperature
                        tmp_raw := analogValues[tmp_analogLower + (tmp_i - tmp_channelsLower)];
                        channels[tmp_i].outputValue := TO_REAL(tmp_raw) / 10.0;
                        channels[tmp_i].retVal := 16#0000;

                    2: // Climatic temperature
                        tmp_raw := analogValues[tmp_analogLower + (tmp_i - tmp_channelsLower)];
                        channels[tmp_i].outputValue := TO_REAL(tmp_raw) / 100.0;
                        channels[tmp_i].retVal := 16#0000;

                    ELSE
                        channels[tmp_i].retVal := 16#8001;
                END_CASE;
            END_IF;
        END_IF;

        tmp_i := tmp_i + 1;
    END_WHILE;

END_FUNCTION_BLOCK

(* ---- public-medium-02.raw_candidate_01.st ---- *)
FUNCTION_BLOCK AnalogBatchProcessing
VAR_INPUT
    count : DINT;
END_VAR
VAR_IN_OUT
    analogValues : ARRAY[*] OF INT;
    channels     : ARRAY[*] OF ST_AnalogChannel;
END_VAR
VAR
    tmp_i         : DINT;
    tmp_rawMin    : REAL;
    tmp_rawMax    : REAL;
    tmp_rawRange  : REAL;
    tmp_engRange  : REAL;
    tmp_raw       : INT;
    tmp_analogVal : REAL;
END_VAR
(* CONTRACT_RULES [] *)
(* ENGINEERING_CONTRACT
 * Activation:       Each scan processes up to 'count' channels sequentially.
 * Retention:        retVal and outputValue are overwritten each scan; no latching.
 * Explicit Reset:   None specified; outputs refresh every scan.
 * Same-scan Priority: Sequential ordinal processing; first failure does not halt loop.
 * Units/Boundaries:
 *   - PUB001: count is caller-supplied bound selector; arrays use their own lower bounds.
 *   - PUB002: measuringMode 0=linear (bipolar/unipolar), 1=std temp (÷10), 2=climatic (÷100).
 *   - PUB003: Linear scaling uses full-scale raw range; output = loLIM + ratio*(hiLIM-loLIM).
 *   - PUB004: RetVal 16#8001 on invalid measuringMode; 16#8002 on hiLIM<=loLIM.
 *   - PUB005: OutputValue written only on successful conversion; retVal set on error.
 *   - PUB006: Disabled channels (enable=FALSE) are skipped without modifying retVal/outputValue.
 *   - PUB007: All arithmetic uses REAL; explicit conversions applied to raw INT operands.
 *   - PUB008: No delay, no edge detection, no state machine; pure per-scan calculation.
 *)

    tmp_i := LOWER_BOUND(analogValues, 1);

    WHILE tmp_i < LOWER_BOUND(analogValues, 1) + count DO
        IF channels[tmp_i].enable THEN
            IF channels[tmp_i].hiLIM <= channels[tmp_i].loLIM THEN
                channels[tmp_i].retVal := 16#8002;
            ELSE
                CASE channels[tmp_i].measuringMode OF
                    0: // Non-temperature linear scaling
                        tmp_raw := analogValues[tmp_i];
                        tmp_analogVal := TO_REAL(tmp_raw);

                        IF channels[tmp_i].bipolar THEN
                            tmp_rawMin := TO_REAL(-27648);
                            tmp_rawMax := TO_REAL(27648);
                        ELSE
                            tmp_rawMin := TO_REAL(0);
                            tmp_rawMax := TO_REAL(27648);
                        END_IF;

                        tmp_rawRange := tmp_rawMax - tmp_rawMin;
                        tmp_engRange := channels[tmp_i].hiLIM - channels[tmp_i].loLIM;

                        channels[tmp_i].outputValue := channels[tmp_i].loLIM +
                            ((tmp_analogVal - tmp_rawMin) / tmp_rawRange) * tmp_engRange;
                        channels[tmp_i].retVal := 16#0000;

                    1: // Standard temperature
                        tmp_raw := analogValues[tmp_i];
                        channels[tmp_i].outputValue := TO_REAL(tmp_raw) / 10.0;
                        channels[tmp_i].retVal := 16#0000;

                    2: // Climatic temperature
                        tmp_raw := analogValues[tmp_i];
                        channels[tmp_i].outputValue := TO_REAL(tmp_raw) / 100.0;
                        channels[tmp_i].retVal := 16#0000;

                    ELSE
                        channels[tmp_i].retVal := 16#8001;
                END_CASE;
            END_IF;
        END_IF;

        tmp_i := tmp_i + 1;
    END_WHILE;

END_FUNCTION_BLOCK

(* ---- public-medium-02.raw_candidate_02.st ---- *)
TYPE ST_AnalogChannel :
STRUCT
    enable        : BOOL;
    hiLIM         : REAL;
    loLIM         : REAL;
    bipolar       : BOOL;
    measuringMode : INT;
    retVal        : WORD;
    outputValue   : REAL;
END_STRUCT
END_TYPE

FUNCTION_BLOCK AnalogBatchProcessing
VAR_INPUT
    count : DINT;
END_VAR
VAR_IN_OUT
    analogValues : ARRAY[*] OF INT;
    channels     : ARRAY[*] OF ST_AnalogChannel;
END_VAR
VAR
    tmp_i         : DINT;
    tmp_rawMin    : REAL;
    tmp_rawMax    : REAL;
    tmp_rawRange  : REAL;
    tmp_engRange  : REAL;
    tmp_raw       : INT;
    tmp_analogVal : REAL;
END_VAR
(* CONTRACT_RULES [] *)
(* ENGINEERING_CONTRACT
 * Activation:       Each scan processes up to 'count' channels sequentially.
 * Retention:        retVal and outputValue are overwritten each scan; no latching.
 * Explicit Reset:   None specified; outputs refresh every scan.
 * Same-scan Priority: Sequential ordinal processing; first failure does not halt loop.
 * Units/Boundaries:
 *   - PUB001: count is caller-supplied bound selector; arrays use their own lower bounds.
 *   - PUB002: measuringMode 0=linear (bipolar/unipolar), 1=std temp (÷10), 2=climatic (÷100).
 *   - PUB003: Linear scaling uses full-scale raw range; output = loLIM + ratio*(hiLIM-loLIM).
 *   - PUB004: RetVal 16#8001 on invalid measuringMode; 16#8002 on hiLIM<=loLIM.
 *   - PUB005: OutputValue written only on successful conversion; retVal set on error.
 *   - PUB006: Disabled channels (enable=FALSE) are skipped without modifying retVal/outputValue.
 *   - PUB007: All arithmetic uses REAL; explicit conversions applied to raw INT operands.
 *   - PUB008: No delay, no edge detection, no state machine; pure per-scan calculation.
 *)

    tmp_i := LOWER_BOUND(analogValues, 1);

    WHILE tmp_i < LOWER_BOUND(analogValues, 1) + count DO
        IF channels[tmp_i].enable THEN
            IF channels[tmp_i].hiLIM <= channels[tmp_i].loLIM THEN
                channels[tmp_i].retVal := 16#8002;
            ELSE
                CASE channels[tmp_i].measuringMode OF
                    0: // Non-temperature linear scaling
                        tmp_raw := analogValues[tmp_i];
                        tmp_analogVal := TO_REAL(tmp_raw);

                        IF channels[tmp_i].bipolar THEN
                            tmp_rawMin := TO_REAL(-27648);
                            tmp_rawMax := TO_REAL(27648);
                        ELSE
                            tmp_rawMin := TO_REAL(0);
                            tmp_rawMax := TO_REAL(27648);
                        END_IF;

                        tmp_rawRange := tmp_rawMax - tmp_rawMin;
                        tmp_engRange := channels[tmp_i].hiLIM - channels[tmp_i].loLIM;

                        channels[tmp_i].outputValue := channels[tmp_i].loLIM +
                            ((tmp_analogVal - tmp_rawMin) / tmp_rawRange) * tmp_engRange;
                        channels[tmp_i].retVal := 16#0000;

                    1: // Standard temperature
                        tmp_raw := analogValues[tmp_i];
                        channels[tmp_i].outputValue := TO_REAL(tmp_raw) / 10.0;
                        channels[tmp_i].retVal := 16#0000;

                    2: // Climatic temperature
                        tmp_raw := analogValues[tmp_i];
                        channels[tmp_i].outputValue := TO_REAL(tmp_raw) / 100.0;
                        channels[tmp_i].retVal := 16#0000;

                    ELSE
                        channels[tmp_i].retVal := 16#8001;
                END_CASE;
            END_IF;
        END_IF;

        tmp_i := tmp_i + 1;
    END_WHILE;

END_FUNCTION_BLOCK

(* ---- public-medium-02.raw_candidate_03.st ---- *)
TYPE ST_AnalogChannel :
STRUCT
    enable        : BOOL;
    hiLIM         : REAL;
    loLIM         : REAL;
    bipolar       : BOOL;
    measuringMode : INT;
    retVal        : WORD;
    outputValue   : REAL;
END_STRUCT
END_TYPE;

FUNCTION_BLOCK AnalogBatchProcessing
VAR_INPUT
    count : DINT;
END_VAR
VAR_IN_OUT
    analogValues : ARRAY[*] OF INT;
    channels     : ARRAY[*] OF ST_AnalogChannel;
END_VAR
VAR
    tmp_i             : DINT;
    tmp_channelsLower : DINT;
    tmp_analogLower   : DINT;
    tmp_rawMin        : REAL;
    tmp_rawMax        : REAL;
    tmp_rawRange      : REAL;
    tmp_engRange      : REAL;
    tmp_raw           : INT;
    tmp_analogVal     : REAL;
END_VAR
(* CONTRACT_RULES [] *)
(* ENGINEERING_CONTRACT
 * Activation:       Each scan processes up to 'count' channels sequentially.
 * Retention:        retVal and outputValue are overwritten each scan; no latching.
 * Explicit Reset:   None specified; outputs refresh every scan.
 * Same-scan Priority: Sequential ordinal processing; first failure does not halt loop.
 * Units/Boundaries:
 *   - PUB001: count is caller-supplied bound selector; arrays use their own lower bounds.
 *   - PUB002: measuringMode 0=linear (bipolar/unipolar), 1=std temp (÷10), 2=climatic (÷100).
 *   - PUB003: Linear scaling uses full-scale raw range; output = loLIM + ratio*(hiLIM-loLIM).
 *   - PUB004: RetVal 16#8001 on invalid measuringMode; 16#8002 on hiLIM<=loLIM.
 *   - PUB005: OutputValue written only on successful conversion; retVal set on error.
 *   - PUB006: Disabled channels (enable=FALSE) are skipped without modifying retVal/outputValue.
 *   - PUB007: All arithmetic uses REAL; explicit conversions applied to raw INT operands.
 *   - PUB008: No delay, no edge detection, no state machine; pure per-scan calculation.
 *)

    tmp_channelsLower := LOWER_BOUND(channels, 1);
    tmp_analogLower   := LOWER_BOUND(analogValues, 1);
    tmp_i := tmp_channelsLower;

    WHILE tmp_i < tmp_channelsLower + count DO
        IF channels[tmp_i].enable THEN
            IF channels[tmp_i].hiLIM <= channels[tmp_i].loLIM THEN
                channels[tmp_i].retVal := 16#8002;
            ELSE
                CASE channels[tmp_i].measuringMode OF
                    0: // Non-temperature linear scaling
                        tmp_raw := analogValues[tmp_analogLower + (tmp_i - tmp_channelsLower)];
                        tmp_analogVal := TO_REAL(tmp_raw);

                        IF channels[tmp_i].bipolar THEN
                            tmp_rawMin := TO_REAL(-27648);
                            tmp_rawMax := TO_REAL(27648);
                        ELSE
                            tmp_rawMin := TO_REAL(0);
                            tmp_rawMax := TO_REAL(27648);
                        END_IF;

                        tmp_rawRange := tmp_rawMax - tmp_rawMin;
                        tmp_engRange := channels[tmp_i].hiLIM - channels[tmp_i].loLIM;

                        channels[tmp_i].outputValue := channels[tmp_i].loLIM +
                            ((tmp_analogVal - tmp_rawMin) / tmp_rawRange) * tmp_engRange;
                        channels[tmp_i].retVal := 16#0000;

                    1: // Standard temperature
                        tmp_raw := analogValues[tmp_analogLower + (tmp_i - tmp_channelsLower)];
                        channels[tmp_i].outputValue := TO_REAL(tmp_raw) / 10.0;
                        channels[tmp_i].retVal := 16#0000;

                    2: // Climatic temperature
                        tmp_raw := analogValues[tmp_analogLower + (tmp_i - tmp_channelsLower)];
                        channels[tmp_i].outputValue := TO_REAL(tmp_raw) / 100.0;
                        channels[tmp_i].retVal := 16#0000;

                    ELSE
                        channels[tmp_i].retVal := 16#8001;
                END_CASE;
            END_IF;
        END_IF;

        tmp_i := tmp_i + 1;
    END_WHILE;

END_FUNCTION_BLOCK

(* ---- public-medium-03.candidate_01.st ---- *)
(*
ENGINEERING_CONTRACT
================================================================================
Output State Summary:
- average:     ACTIVATION on cyclicExecution=TRUE OR rising trigger edge | RETAIN between updates
- windowSizeReached: RETAIN | FALSE until sampleCount>=windowSize | reset clears to FALSE
- error:       RETAIN | set TRUE on windowSize outside [1,100] | reset clears to FALSE
- status:      RETAIN | 16#0000=success, 16#8200=windowSize error | reset clears to 16#0000

Scan Priority (same-scan):
- cyclicExecution=TRUE → add value and exit; trigger ignored (PUB001/PUB002 priority)
- cyclicExecution=FALSE AND trigger rising edge → add value (PUB002)

Reset Behavior (PUB005):
- reset=TRUE → clear all state, set status=16#0000, error=FALSE; no output update same scan
- reset is level-triggered; next scan after reset=FALSE resumes normal operation

Boundary Constraints:
- windowSize: [1,100] inclusive (PUB003)
- average = sum / windowSize when sampleCount>=windowSize, else sum/sampleCount
- Division guard: MAX(1,sampleCount) prevents zero-divide on first value
================================================================================
*)

(* CONTRACT_RULES [] *)

FUNCTION_BLOCK FB_MovingAverage
VAR_INPUT
    cyclicExecution : BOOL;
    trigger : BOOL;
    value : LREAL;
    windowSize : INT;
    reset : BOOL;
END_VAR

VAR_OUTPUT
    average : LREAL := 0.0;
    windowSizeReached : BOOL := FALSE;
    error : BOOL := FALSE;
    status : WORD := 16#0000;
END_VAR

VAR
    dataBuffer : ARRAY[1..100] OF LREAL;
    currentIndex : INT := 0;
    sampleCount : INT := 0;
    sum : LREAL := 0.0;
    prevTrigger : BOOL := FALSE;
END_VAR

METHOD PRIVATE AddValueAndUpdateAverage : BOOL
VAR
    oldestValue : LREAL;
END_VAR

    oldestValue := 0.0;

    IF sampleCount >= windowSize THEN
        oldestValue := dataBuffer[currentIndex];
    END_IF;

    dataBuffer[currentIndex] := value;
    sum := sum + value - oldestValue;

    currentIndex := currentIndex + 1;
    IF currentIndex > windowSize THEN
        currentIndex := 1;
    END_IF;

    IF sampleCount < windowSize THEN
        sampleCount := sampleCount + 1;
    END_IF;

    windowSizeReached := (sampleCount >= windowSize);

    average := sum / TO_LREAL(MAX(1, sampleCount));

    AddValueAndUpdateAverage := TRUE;
END_METHOD

IF reset THEN
    currentIndex := 0;
    sampleCount := 0;
    sum := 0.0;
    windowSizeReached := FALSE;
    error := FALSE;
    status := 16#0000;
    average := 0.0;
    prevTrigger := trigger;
    RETURN;
END_IF;

IF windowSize < 1 OR windowSize > 100 THEN
    error := TRUE;
    status := 16#8200;
    prevTrigger := trigger;
    RETURN;
END_IF;

error := FALSE;
status := 16#0000;

IF cyclicExecution THEN
    AddValueAndUpdateAverage();
ELSIF trigger AND NOT prevTrigger THEN
    AddValueAndUpdateAverage();
END_IF;

prevTrigger := trigger;
END_FUNCTION_BLOCK

(* ---- public-medium-03.candidate_02.st ---- *)
(* ENGINEERING_CONTRACT
================================================================================
Output State Summary:
- average:     ACTIVATION on cyclicExecution=TRUE OR rising trigger edge | RETAIN between updates
- windowSizeReached: RETAIN | FALSE until sampleCount>=windowSize | reset clears to FALSE
- error:       RETAIN | set TRUE on windowSize outside [1,100] | reset clears to FALSE
- status:      RETAIN | 16#0000=success, 16#8200=windowSize error | reset clears to 16#0000

Scan Priority (same-scan):
- cyclicExecution=TRUE → add value and exit; trigger ignored (PUB001/PUB002 priority)
- cyclicExecution=FALSE AND trigger rising edge → add value (PUB002)

Reset Behavior (PUB005):
- reset=TRUE → clear all state, set status=16#0000, error=FALSE; no output update same scan
- reset is level-triggered; next scan after reset=FALSE resumes normal operation

Boundary Constraints:
- windowSize: [1,100] inclusive (PUB003)
- average = sum / windowSize when sampleCount>=windowSize, else sum/sampleCount
- Division guard: MAX(1,sampleCount) prevents zero-divide on first value
================================================================================
*)

(* CONTRACT_RULES [] *)

FUNCTION_BLOCK FB_MovingAverage
VAR_INPUT
    cyclicExecution : BOOL;
    trigger : BOOL;
    value : LREAL;
    windowSize : INT;
    reset : BOOL;
END_VAR

VAR_OUTPUT
    average : LREAL := 0.0;
    windowSizeReached : BOOL := FALSE;
    error : BOOL := FALSE;
    status : WORD := 16#0000;
END_VAR

VAR
    dataBuffer : ARRAY[1..100] OF LREAL;
    currentIndex : INT := 0;
    sampleCount : INT := 0;
    sum : LREAL := 0.0;
    prevTrigger : BOOL := FALSE;
END_VAR

VAR
    tmpAddValue : BOOL;
    tmpOldestValue : LREAL;
END_VAR

tmpAddValue := FALSE;

IF reset THEN
    currentIndex := 0;
    sampleCount := 0;
    sum := 0.0;
    windowSizeReached := FALSE;
    error := FALSE;
    status := 16#0000;
    average := 0.0;
    prevTrigger := trigger;
    RETURN;
END_IF;

IF windowSize < 1 OR windowSize > 100 THEN
    error := TRUE;
    status := 16#8200;
    prevTrigger := trigger;
    RETURN;
END_IF;

error := FALSE;
status := 16#0000;

IF cyclicExecution THEN
    tmpAddValue := TRUE;
ELSIF trigger AND NOT prevTrigger THEN
    tmpAddValue := TRUE;
END_IF;

IF tmpAddValue THEN
    tmpOldestValue := 0.0;

    IF sampleCount >= windowSize THEN
        tmpOldestValue := dataBuffer[currentIndex];
    END_IF;

    dataBuffer[currentIndex] := value;
    sum := sum + value - tmpOldestValue;

    currentIndex := currentIndex + 1;
    IF currentIndex > windowSize THEN
        currentIndex := 1;
    END_IF;

    IF sampleCount < windowSize THEN
        sampleCount := sampleCount + 1;
    END_IF;

    windowSizeReached := (sampleCount >= windowSize);

    average := sum / TO_LREAL(MAX(1, sampleCount));
END_IF;

prevTrigger := trigger;
END_FUNCTION_BLOCK

(* ---- public-medium-03.candidate_03.st ---- *)
(* ENGINEERING_CONTRACT
================================================================================
Output State Summary:
- average:     ACTIVATION on cyclicExecution=TRUE OR rising trigger edge | RETAIN
- windowSizeReached: RETAIN | FALSE until sampleCount>=windowSize | reset clears
- error:       RETAIN | set TRUE on windowSize outside [1,100] | reset clears
- status:      RETAIN | 16#0000=success, 16#8200=windowSize error | reset clears

Scan Priority (same-scan):
- cyclicExecution=TRUE → add value (trigger ignored) [PUB001/PUB002 priority]
- cyclicExecution=FALSE AND trigger rising edge → add value [PUB002]

Reset Behavior (PUB005):
- reset=TRUE → clear all state, set status=16#0000, exit immediately

Boundary Constraints (PUB003):
- windowSize: [1,100] inclusive
- average = sum / MIN(windowSize, sampleCount) when full, else sum/sampleCount
- Division guard: MAX(1,sampleCount) prevents zero-divide [PUB001]
================================================================================
*)

(* CONTRACT_RULES [] *)

FUNCTION_BLOCK FB_MovingAverage
VAR_INPUT
    cyclicExecution : BOOL;
    trigger : BOOL;
    value : LREAL;
    windowSize : INT;
    reset : BOOL;
END_VAR

VAR_OUTPUT
    average : LREAL := 0.0;
    windowSizeReached : BOOL := FALSE;
    error : BOOL := FALSE;
    status : WORD := 16#0000;
END_VAR

VAR
    dataBuffer : ARRAY[1..100] OF LREAL;
    currentIndex : INT := 0;
    sampleCount : INT := 0;
    sum : LREAL := 0.0;
    prevTrigger : BOOL := FALSE;
    evictIndex : INT := 1;
END_VAR

VAR
    tmpAddValue : BOOL;
    tmpOldestValue : LREAL;
END_VAR

tmpAddValue := FALSE;

IF reset THEN
    currentIndex := 0;
    sampleCount := 0;
    sum := 0.0;
    windowSizeReached := FALSE;
    error := FALSE;
    status := 16#0000;
    average := 0.0;
    prevTrigger := trigger;
    RETURN;
END_IF;

IF windowSize < 1 OR windowSize > 100 THEN
    error := TRUE;
    status := 16#8200;
    prevTrigger := trigger;
    RETURN;
END_IF;

error := FALSE;
status := 16#0000;

IF cyclicExecution THEN
    tmpAddValue := TRUE;
ELSIF trigger AND NOT prevTrigger THEN
    tmpAddValue := TRUE;
END_IF;

IF tmpAddValue THEN
    tmpOldestValue := 0.0;

    IF sampleCount >= windowSize THEN
        tmpOldestValue := dataBuffer[evictIndex];
        evictIndex := evictIndex + 1;
        IF evictIndex > windowSize THEN
            evictIndex := 1;
        END_IF;
    END_IF;

    currentIndex := currentIndex + 1;
    IF currentIndex > windowSize THEN
        currentIndex := 1;
    END_IF;

    dataBuffer[currentIndex] := value;
    sum := sum + value - tmpOldestValue;

    IF sampleCount < windowSize THEN
        sampleCount := sampleCount + 1;
    END_IF;

    windowSizeReached := (sampleCount >= windowSize);

    average := sum / TO_LREAL(MAX(1, sampleCount));
END_IF;

prevTrigger := trigger;
END_FUNCTION_BLOCK

(* ---- public-medium-03.candidate_04.st ---- *)
(* ENGINEERING_CONTRACT
================================================================================
Output State Summary:
- average:     ACTIVATION on cyclicExecution=TRUE OR rising trigger edge | RETAIN
- windowSizeReached: RETAIN | FALSE until sampleCount>=windowSize | reset clears
- error:       RETAIN | set TRUE on windowSize outside [1,100] | reset clears
- status:      RETAIN | 16#0000=success, 16#8200=windowSize error | reset clears

Scan Priority (same-scan):
- cyclicExecution=TRUE → add value (trigger ignored) [PUB001/PUB002 priority]
- cyclicExecution=FALSE AND trigger rising edge → add value [PUB002]

Reset Behavior (PUB005):
- reset=TRUE → clear all state, set status=16#0000, exit immediately

Boundary Constraints (PUB003):
- windowSize: [1,100] inclusive
- average = sum / MIN(windowSize, sampleCount) when full, else sum/sampleCount
- Division guard: MAX(1,sampleCount) prevents zero-divide [PUB001]
- Window shrink: reset sampleCount and sum to force clean restart [replay fix]
================================================================================
*)

(* CONTRACT_RULES [] *)

FUNCTION_BLOCK FB_MovingAverage
VAR_INPUT
    cyclicExecution : BOOL;
    trigger : BOOL;
    value : LREAL;
    windowSize : INT;
    reset : BOOL;
END_VAR

VAR_OUTPUT
    average : LREAL := 0.0;
    windowSizeReached : BOOL := FALSE;
    error : BOOL := FALSE;
    status : WORD := 16#0000;
END_VAR

VAR
    dataBuffer : ARRAY[1..100] OF LREAL;
    currentIndex : INT := 0;
    sampleCount : INT := 0;
    sum : LREAL := 0.0;
    prevTrigger : BOOL := FALSE;
    evictIndex : INT := 1;
    prevWindowSize : INT := 0;
END_VAR

VAR
    tmpAddValue : BOOL;
    tmpOldestValue : LREAL;
    tmp_WindowSizeChanged : BOOL;
END_VAR

tmpAddValue := FALSE;
tmp_WindowSizeChanged := FALSE;

IF reset THEN
    currentIndex := 0;
    sampleCount := 0;
    sum := 0.0;
    windowSizeReached := FALSE;
    error := FALSE;
    status := 16#0000;
    average := 0.0;
    prevTrigger := trigger;
    prevWindowSize := windowSize;
    RETURN;
END_IF;

IF windowSize < 1 OR windowSize > 100 THEN
    error := TRUE;
    status := 16#8200;
    prevTrigger := trigger;
    prevWindowSize := windowSize;
    RETURN;
END_IF;

error := FALSE;
status := 16#0000;

IF windowSize < prevWindowSize AND sampleCount > windowSize THEN
    tmp_WindowSizeChanged := TRUE;
    sampleCount := 0;
    sum := 0.0;
    currentIndex := 0;
    evictIndex := 1;
END_IF;

IF cyclicExecution THEN
    tmpAddValue := TRUE;
ELSIF trigger AND NOT prevTrigger THEN
    tmpAddValue := TRUE;
END_IF;

IF tmpAddValue THEN
    tmpOldestValue := 0.0;

    IF sampleCount >= windowSize THEN
        tmpOldestValue := dataBuffer[evictIndex];
        evictIndex := evictIndex + 1;
        IF evictIndex > windowSize THEN
            evictIndex := 1;
        END_IF;
    END_IF;

    currentIndex := currentIndex + 1;
    IF currentIndex > windowSize THEN
        currentIndex := 1;
    END_IF;

    dataBuffer[currentIndex] := value;
    sum := sum + value - tmpOldestValue;

    IF sampleCount < windowSize THEN
        sampleCount := sampleCount + 1;
    END_IF;

    windowSizeReached := (sampleCount >= windowSize);

    average := sum / TO_LREAL(MAX(1, sampleCount));
END_IF;

prevTrigger := trigger;
prevWindowSize := windowSize;
END_FUNCTION_BLOCK

(* ---- public-medium-03.raw_candidate_01.st ---- *)
(*
ENGINEERING_CONTRACT
================================================================================
Output State Summary:
- average:     ACTIVATION on cyclicExecution=TRUE OR rising trigger edge | RETAIN between updates
- windowSizeReached: RETAIN | FALSE until sampleCount>=windowSize | reset clears to FALSE
- error:       RETAIN | set TRUE on windowSize outside [1,100] | reset clears to FALSE
- status:      RETAIN | 16#0000=success, 16#8200=windowSize error | reset clears to 16#0000

Scan Priority (same-scan):
- cyclicExecution=TRUE → add value and exit; trigger ignored (PUB001/PUB002 priority)
- cyclicExecution=FALSE AND trigger rising edge → add value (PUB002)

Reset Behavior (PUB005):
- reset=TRUE → clear all state, set status=16#0000, error=FALSE; no output update same scan
- reset is level-triggered; next scan after reset=FALSE resumes normal operation

Boundary Constraints:
- windowSize: [1,100] inclusive (PUB003)
- average = sum / windowSize when sampleCount>=windowSize, else sum/sampleCount
- Division guard: MAX(1,sampleCount) prevents zero-divide on first value
================================================================================
*)

(* CONTRACT_RULES [] *)

FUNCTION_BLOCK FB_MovingAverage
VAR_INPUT
    cyclicExecution : BOOL;
    trigger : BOOL;
    value : LREAL;
    windowSize : INT;
    reset : BOOL;
END_VAR

VAR_OUTPUT
    average : LREAL := 0.0;
    windowSizeReached : BOOL := FALSE;
    error : BOOL := FALSE;
    status : WORD := 16#0000;
END_VAR

VAR
    dataBuffer : ARRAY[1..100] OF LREAL;
    currentIndex : INT := 0;
    sampleCount : INT := 0;
    sum : LREAL := 0.0;
    prevTrigger : BOOL := FALSE;
END_VAR

METHOD PRIVATE AddValueAndUpdateAverage : BOOL
VAR
    oldestValue : LREAL;
END_VAR

    oldestValue := 0.0;

    IF sampleCount >= windowSize THEN
        oldestValue := dataBuffer[currentIndex];
    END_IF;

    dataBuffer[currentIndex] := value;
    sum := sum + value - oldestValue;

    currentIndex := currentIndex + 1;
    IF currentIndex > windowSize THEN
        currentIndex := 1;
    END_IF;

    IF sampleCount < windowSize THEN
        sampleCount := sampleCount + 1;
    END_IF;

    windowSizeReached := (sampleCount >= windowSize);

    average := sum / TO_LREAL(MAX(1, sampleCount));

    AddValueAndUpdateAverage := TRUE;
END_METHOD

IF reset THEN
    currentIndex := 0;
    sampleCount := 0;
    sum := 0.0;
    windowSizeReached := FALSE;
    error := FALSE;
    status := 16#0000;
    average := 0.0;
    prevTrigger := trigger;
    RETURN;
END_IF;

IF windowSize < 1 OR windowSize > 100 THEN
    error := TRUE;
    status := 16#8200;
    prevTrigger := trigger;
    RETURN;
END_IF;

error := FALSE;
status := 16#0000;

IF cyclicExecution THEN
    AddValueAndUpdateAverage();
ELSIF trigger AND NOT prevTrigger THEN
    AddValueAndUpdateAverage();
END_IF;

prevTrigger := trigger;
END_FUNCTION_BLOCK

(* ---- public-medium-03.raw_candidate_02.st ---- *)
(* ENGINEERING_CONTRACT
================================================================================
Output State Summary:
- average:     ACTIVATION on cyclicExecution=TRUE OR rising trigger edge | RETAIN between updates
- windowSizeReached: RETAIN | FALSE until sampleCount>=windowSize | reset clears to FALSE
- error:       RETAIN | set TRUE on windowSize outside [1,100] | reset clears to FALSE
- status:      RETAIN | 16#0000=success, 16#8200=windowSize error | reset clears to 16#0000

Scan Priority (same-scan):
- cyclicExecution=TRUE → add value and exit; trigger ignored (PUB001/PUB002 priority)
- cyclicExecution=FALSE AND trigger rising edge → add value (PUB002)

Reset Behavior (PUB005):
- reset=TRUE → clear all state, set status=16#0000, error=FALSE; no output update same scan
- reset is level-triggered; next scan after reset=FALSE resumes normal operation

Boundary Constraints:
- windowSize: [1,100] inclusive (PUB003)
- average = sum / windowSize when sampleCount>=windowSize, else sum/sampleCount
- Division guard: MAX(1,sampleCount) prevents zero-divide on first value
================================================================================
*)

(* CONTRACT_RULES [] *)

FUNCTION_BLOCK FB_MovingAverage
VAR_INPUT
    cyclicExecution : BOOL;
    trigger : BOOL;
    value : LREAL;
    windowSize : INT;
    reset : BOOL;
END_VAR

VAR_OUTPUT
    average : LREAL := 0.0;
    windowSizeReached : BOOL := FALSE;
    error : BOOL := FALSE;
    status : WORD := 16#0000;
END_VAR

VAR
    dataBuffer : ARRAY[1..100] OF LREAL;
    currentIndex : INT := 0;
    sampleCount : INT := 0;
    sum : LREAL := 0.0;
    prevTrigger : BOOL := FALSE;
END_VAR

VAR
    tmpAddValue : BOOL;
    tmpOldestValue : LREAL;
END_VAR

tmpAddValue := FALSE;

IF reset THEN
    currentIndex := 0;
    sampleCount := 0;
    sum := 0.0;
    windowSizeReached := FALSE;
    error := FALSE;
    status := 16#0000;
    average := 0.0;
    prevTrigger := trigger;
    RETURN;
END_IF;

IF windowSize < 1 OR windowSize > 100 THEN
    error := TRUE;
    status := 16#8200;
    prevTrigger := trigger;
    RETURN;
END_IF;

error := FALSE;
status := 16#0000;

IF cyclicExecution THEN
    tmpAddValue := TRUE;
ELSIF trigger AND NOT prevTrigger THEN
    tmpAddValue := TRUE;
END_IF;

IF tmpAddValue THEN
    tmpOldestValue := 0.0;

    IF sampleCount >= windowSize THEN
        tmpOldestValue := dataBuffer[currentIndex];
    END_IF;

    dataBuffer[currentIndex] := value;
    sum := sum + value - tmpOldestValue;

    currentIndex := currentIndex + 1;
    IF currentIndex > windowSize THEN
        currentIndex := 1;
    END_IF;

    IF sampleCount < windowSize THEN
        sampleCount := sampleCount + 1;
    END_IF;

    windowSizeReached := (sampleCount >= windowSize);

    average := sum / TO_LREAL(MAX(1, sampleCount));
END_IF;

prevTrigger := trigger;
END_FUNCTION_BLOCK

(* ---- public-medium-03.raw_candidate_03.st ---- *)
(* ENGINEERING_CONTRACT
================================================================================
Output State Summary:
- average:     ACTIVATION on cyclicExecution=TRUE OR rising trigger edge | RETAIN
- windowSizeReached: RETAIN | FALSE until sampleCount>=windowSize | reset clears
- error:       RETAIN | set TRUE on windowSize outside [1,100] | reset clears
- status:      RETAIN | 16#0000=success, 16#8200=windowSize error | reset clears

Scan Priority (same-scan):
- cyclicExecution=TRUE → add value (trigger ignored) [PUB001/PUB002 priority]
- cyclicExecution=FALSE AND trigger rising edge → add value [PUB002]

Reset Behavior (PUB005):
- reset=TRUE → clear all state, set status=16#0000, exit immediately

Boundary Constraints (PUB003):
- windowSize: [1,100] inclusive
- average = sum / MIN(windowSize, sampleCount) when full, else sum/sampleCount
- Division guard: MAX(1,sampleCount) prevents zero-divide [PUB001]
================================================================================
*)

(* CONTRACT_RULES [] *)

FUNCTION_BLOCK FB_MovingAverage
VAR_INPUT
    cyclicExecution : BOOL;
    trigger : BOOL;
    value : LREAL;
    windowSize : INT;
    reset : BOOL;
END_VAR

VAR_OUTPUT
    average : LREAL := 0.0;
    windowSizeReached : BOOL := FALSE;
    error : BOOL := FALSE;
    status : WORD := 16#0000;
END_VAR

VAR
    dataBuffer : ARRAY[1..100] OF LREAL;
    currentIndex : INT := 0;
    sampleCount : INT := 0;
    sum : LREAL := 0.0;
    prevTrigger : BOOL := FALSE;
    evictIndex : INT := 1;
END_VAR

VAR
    tmpAddValue : BOOL;
    tmpOldestValue : LREAL;
END_VAR

tmpAddValue := FALSE;

IF reset THEN
    currentIndex := 0;
    sampleCount := 0;
    sum := 0.0;
    windowSizeReached := FALSE;
    error := FALSE;
    status := 16#0000;
    average := 0.0;
    prevTrigger := trigger;
    RETURN;
END_IF;

IF windowSize < 1 OR windowSize > 100 THEN
    error := TRUE;
    status := 16#8200;
    prevTrigger := trigger;
    RETURN;
END_IF;

error := FALSE;
status := 16#0000;

IF cyclicExecution THEN
    tmpAddValue := TRUE;
ELSIF trigger AND NOT prevTrigger THEN
    tmpAddValue := TRUE;
END_IF;

IF tmpAddValue THEN
    tmpOldestValue := 0.0;

    IF sampleCount >= windowSize THEN
        tmpOldestValue := dataBuffer[evictIndex];
        evictIndex := evictIndex + 1;
        IF evictIndex > windowSize THEN
            evictIndex := 1;
        END_IF;
    END_IF;

    currentIndex := currentIndex + 1;
    IF currentIndex > windowSize THEN
        currentIndex := 1;
    END_IF;

    dataBuffer[currentIndex] := value;
    sum := sum + value - tmpOldestValue;

    IF sampleCount < windowSize THEN
        sampleCount := sampleCount + 1;
    END_IF;

    windowSizeReached := (sampleCount >= windowSize);

    average := sum / TO_LREAL(MAX(1, sampleCount));
END_IF;

prevTrigger := trigger;
END_FUNCTION_BLOCK

(* ---- public-medium-03.raw_candidate_04.st ---- *)
(* ENGINEERING_CONTRACT
================================================================================
Output State Summary:
- average:     ACTIVATION on cyclicExecution=TRUE OR rising trigger edge | RETAIN
- windowSizeReached: RETAIN | FALSE until sampleCount>=windowSize | reset clears
- error:       RETAIN | set TRUE on windowSize outside [1,100] | reset clears
- status:      RETAIN | 16#0000=success, 16#8200=windowSize error | reset clears

Scan Priority (same-scan):
- cyclicExecution=TRUE → add value (trigger ignored) [PUB001/PUB002 priority]
- cyclicExecution=FALSE AND trigger rising edge → add value [PUB002]

Reset Behavior (PUB005):
- reset=TRUE → clear all state, set status=16#0000, exit immediately

Boundary Constraints (PUB003):
- windowSize: [1,100] inclusive
- average = sum / MIN(windowSize, sampleCount) when full, else sum/sampleCount
- Division guard: MAX(1,sampleCount) prevents zero-divide [PUB001]
- Window shrink: reset sampleCount and sum to force clean restart [replay fix]
================================================================================
*)

(* CONTRACT_RULES [] *)

FUNCTION_BLOCK FB_MovingAverage
VAR_INPUT
    cyclicExecution : BOOL;
    trigger : BOOL;
    value : LREAL;
    windowSize : INT;
    reset : BOOL;
END_VAR

VAR_OUTPUT
    average : LREAL := 0.0;
    windowSizeReached : BOOL := FALSE;
    error : BOOL := FALSE;
    status : WORD := 16#0000;
END_VAR

VAR
    dataBuffer : ARRAY[1..100] OF LREAL;
    currentIndex : INT := 0;
    sampleCount : INT := 0;
    sum : LREAL := 0.0;
    prevTrigger : BOOL := FALSE;
    evictIndex : INT := 1;
    prevWindowSize : INT := 0;
END_VAR

VAR
    tmpAddValue : BOOL;
    tmpOldestValue : LREAL;
    tmp_WindowSizeChanged : BOOL;
END_VAR

tmpAddValue := FALSE;
tmp_WindowSizeChanged := FALSE;

IF reset THEN
    currentIndex := 0;
    sampleCount := 0;
    sum := 0.0;
    windowSizeReached := FALSE;
    error := FALSE;
    status := 16#0000;
    average := 0.0;
    prevTrigger := trigger;
    prevWindowSize := windowSize;
    RETURN;
END_IF;

IF windowSize < 1 OR windowSize > 100 THEN
    error := TRUE;
    status := 16#8200;
    prevTrigger := trigger;
    prevWindowSize := windowSize;
    RETURN;
END_IF;

error := FALSE;
status := 16#0000;

IF windowSize < prevWindowSize AND sampleCount > windowSize THEN
    tmp_WindowSizeChanged := TRUE;
    sampleCount := 0;
    sum := 0.0;
    currentIndex := 0;
    evictIndex := 1;
END_IF;

IF cyclicExecution THEN
    tmpAddValue := TRUE;
ELSIF trigger AND NOT prevTrigger THEN
    tmpAddValue := TRUE;
END_IF;

IF tmpAddValue THEN
    tmpOldestValue := 0.0;

    IF sampleCount >= windowSize THEN
        tmpOldestValue := dataBuffer[evictIndex];
        evictIndex := evictIndex + 1;
        IF evictIndex > windowSize THEN
            evictIndex := 1;
        END_IF;
    END_IF;

    currentIndex := currentIndex + 1;
    IF currentIndex > windowSize THEN
        currentIndex := 1;
    END_IF;

    dataBuffer[currentIndex] := value;
    sum := sum + value - tmpOldestValue;

    IF sampleCount < windowSize THEN
        sampleCount := sampleCount + 1;
    END_IF;

    windowSizeReached := (sampleCount >= windowSize);

    average := sum / TO_LREAL(MAX(1, sampleCount));
END_IF;

prevTrigger := trigger;
prevWindowSize := windowSize;
END_FUNCTION_BLOCK

(* ---- public-medium-04.candidate_01.st ---- *)
(*
ENGINEERING_CONTRACT:
PUB001: Read TemperatureSensorInput (REAL), display in CurrentTemperature
PUB002: HeaterOutput := TRUE when TemperatureSensorInput < SetTemperature
PUB003: Overheat triggers after >5s continuous HeaterOutput (strict > boundary)
PUB004: Overheat auto-sets HeaterOutput:=FALSE, 3s cooldown before OverheatProtection can clear
PUB005: Sensor fault (<0 OR >100) sets HeaterOutput:=FALSE regardless of temperature
PUB006: Status outputs (CurrentTemperature, SetTempDisplay, HeaterStatus, OverheatProtection) update every scan

Activation: All outputs update every scan (no edge-only behavior)
Retention: OverheatActive retains state across scans until cooldown completes
Reset/Deactivation: OverheatActive resets only after OverheatCooldownTimer.Q (3s elapsed)
Same-scan priority: HeaterOutput finalized BEFORE runtime timer enable is evaluated
Units: TIME/LTIME for timers (TON), REAL for temperatures, BOOL for control/status
*)
FUNCTION_BLOCK FB_TemperatureControl
VAR_INPUT
    TemperatureSensorInput : REAL;
    SetTemperature : REAL;
END_VAR

VAR_OUTPUT
    CurrentTemperature : REAL;
    SetTempDisplay : REAL;
    HeaterStatus : BOOL;
    OverheatProtection : BOOL;
    HeaterOutput : BOOL;
END_VAR

VAR
    HeaterRuntimeTimer : TON;
    OverheatCooldownTimer : TON;
    OverheatActive : BOOL := FALSE;
    SensorFault : BOOL := FALSE;
END_VAR

// Update display outputs
CurrentTemperature := TemperatureSensorInput;
SetTempDisplay := SetTemperature;

// Sensor fault detection: invalid range turns off heater
SensorFault := (TemperatureSensorInput < 0.0) OR (TemperatureSensorInput > 100.0);

// Temperature control logic
IF NOT SensorFault AND NOT OverheatActive THEN
    // Normal operation: heater ON when below setpoint
    IF TemperatureSensorInput < SetTemperature THEN
        HeaterOutput := TRUE;
    ELSE
        HeaterOutput := FALSE;
    END_IF;
ELSE
    // Sensor fault or overheat protection active - heater OFF
    HeaterOutput := FALSE;
END_IF;

// Update heater status display
HeaterStatus := HeaterOutput;

// Runtime timer: tracks continuous heater ON time (resets when heater OFF)
HeaterRuntimeTimer(IN := HeaterOutput, PT := T#5s);

// Overheat detection: >5s continuous heater operation
IF HeaterRuntimeTimer.Q AND NOT OverheatActive THEN
    OverheatActive := TRUE;
    OverheatCooldownTimer(IN := TRUE, PT := T#3s);
END_IF;

// Overheat cooldown: 3s wait before protection can be lifted
IF OverheatActive THEN
    OverheatCooldownTimer(IN := TRUE, PT := T#3s);
    IF OverheatCooldownTimer.Q THEN
        OverheatActive := FALSE;
    END_IF;
END_IF;

// Update overheat protection status
OverheatProtection := OverheatActive;
END_FUNCTION_BLOCK

(* ---- public-medium-04.candidate_02.st ---- *)
(*
ENGINEERING_CONTRACT:
PUB001: TemperatureSensorInput (REAL) -> CurrentTemperature (REAL) every scan
PUB002: HeaterOutput := TRUE when TemperatureSensorInput < SetTemperature (no sensor fault)
PUB003: Overheat triggers when runtime > 5s (strict >), first satisfying tick = 5001ms
PUB004: Overheat sets HeaterOutput:=FALSE, 3s cooldown before OverheatProtection clears
PUB005: Sensor fault (<0 OR >100) sets HeaterOutput:=FALSE regardless of temperature
PUB006: All status outputs (CurrentTemperature, SetTempDisplay, HeaterStatus, OverheatProtection) update every scan
*)
FUNCTION_BLOCK FB_TemperatureControl
VAR_INPUT
    TemperatureSensorInput : REAL;
    SetTemperature         : REAL;
END_VAR

VAR_OUTPUT
    CurrentTemperature : REAL;
    SetTempDisplay      : REAL;
    HeaterStatus        : BOOL;
    OverheatProtection  : BOOL;
    HeaterOutput        : BOOL;
END_VAR

VAR
    HeaterRuntimeTimer   : TON;
    OverheatCooldownTimer: TON;
    OverheatActive       : BOOL := FALSE;
    SensorFault          : BOOL := FALSE;
    Runtimems            : LINT := 0;
END_VAR

SensorFault := (TemperatureSensorInput < 0.0) OR (TemperatureSensorInput > 100.0);

IF NOT SensorFault AND NOT OverheatActive THEN
    IF TemperatureSensorInput < SetTemperature THEN
        HeaterOutput := TRUE;
    ELSE
        HeaterOutput := FALSE;
    END_IF;
ELSE
    HeaterOutput := FALSE;
END_IF;

HeaterRuntimeTimer(IN := FALSE, PT := T#5s);

IF OverheatActive THEN
    IF Runtimems > 5000 THEN
        OverheatActive := TRUE;
    END_IF;
ELSIF HeaterOutput THEN
    Runtimems := Runtimems + TO_LINT(HeaterRuntimeTimer.ET) + 1;
    HeaterRuntimeTimer(IN := TRUE, PT := T#5s);
    IF Runtimems > 5000 THEN
        OverheatActive := TRUE;
        HeaterOutput := FALSE;
    END_IF;
ELSE
    Runtimems := 0;
END_IF;

IF OverheatActive THEN
    OverheatCooldownTimer(IN := TRUE, PT := T#3s);
    IF OverheatCooldownTimer.Q THEN
        OverheatActive := FALSE;
        Runtimems := 0;
    END_IF;
END_IF;

CurrentTemperature := TemperatureSensorInput;
SetTempDisplay := SetTemperature;
HeaterStatus := HeaterOutput;
OverheatProtection := OverheatActive;
END_FUNCTION_BLOCK

(* ---- public-medium-04.candidate_03.st ---- *)
(* CONTRACT_RULES [] *)
FUNCTION_BLOCK FB_TemperatureControl
VAR_INPUT
    TemperatureSensorInput : REAL;
    SetTemperature : REAL;
END_VAR
VAR_OUTPUT
    CurrentTemperature : REAL;
    SetTempDisplay : REAL;
    HeaterStatus : BOOL;
    OverheatProtection : BOOL;
    HeaterOutput : BOOL;
END_VAR
VAR
    HeaterRuntimeTimer : TON;
    OverheatCooldownTimer : TON;
    OverheatActive : BOOL := FALSE;
    SensorFault : BOOL := FALSE;
END_VAR

CurrentTemperature := TemperatureSensorInput;
SetTempDisplay := SetTemperature;
SensorFault := (TemperatureSensorInput < 0.0) OR (TemperatureSensorInput > 100.0);

HeaterRuntimeTimer(IN := (TemperatureSensorInput < SetTemperature) AND NOT SensorFault AND NOT OverheatActive, PT := T#5s);

IF HeaterRuntimeTimer.Q AND NOT OverheatActive THEN
    OverheatActive := TRUE;
    OverheatCooldownTimer(IN := TRUE, PT := T#3s);
END_IF;

IF OverheatActive THEN
    OverheatCooldownTimer(IN := TRUE, PT := T#3s);
    IF OverheatCooldownTimer.Q THEN
        OverheatActive := FALSE;
    END_IF;
END_IF;

IF NOT SensorFault AND NOT OverheatActive THEN
    IF TemperatureSensorInput < SetTemperature THEN
        HeaterOutput := TRUE;
    ELSE
        HeaterOutput := FALSE;
    END_IF;
ELSE
    HeaterOutput := FALSE;
END_IF;

HeaterStatus := HeaterOutput;
OverheatProtection := OverheatActive;
END_FUNCTION_BLOCK
